(* IEC 61131-3 sources: daoli-st-library/DL_Base (part 12) *)

(* ---- FB_DL_EventCounter.st ---- *)
(*==============================================================================
 * 组件名称 (Component)  : FB_DL_EventCounter
 * 所属子库 (Sublibrary) : DL_Base
 * 当前版本 (Version)    : 1.0.1
 * 兼容性   (Platform)   : CODESYS 3.5 / TwinCAT 3 / 汇川 InoProShop / Machine Expert
 *                         仅依赖 Standard.library（R_TRIG），零厂商方言
 * 分类     (Category)   : 信号处理功能块（Function Block · 通用事件计数）
 * 功能简述 (Function)   : 双向事件计数器（DINT 域）。递增/递减脉冲沿独立
 *                         计数、预置装载、高/低阈值比较输出（每拍重算非锁
 *                         存）、回绕/饱和两种越界模式可选；双脉冲同拍抵消
 *                         置信息级、装载覆盖计数置信息级；参数非法故障锁存。
 *                         与 FC_DL_BitCount（位统计）、FB_DL_RuntimeMeter
 *                         （时间累计）职责分离，本块为通用事件计数。
 * 公约遵循 (Convention) : 0.1/R23 事件型，免首扫——计数由脉冲沿驱动，无
 *                         初始化/跟踪同步语义，不设 bInit。
 *                         0.2/R21 bFault 为显式排除信息级码的派生式；故障
 *                         码表逐条标注级别；信息级只进 uErrorId 不进报警链。
 *                         0.7/R15 故障级锁存仅解除路径（bReset 上升沿）清
 *                         码；信息级瞬时型每拍重算。
 *                         0.8 故障码段位 16#0001_xxxx（经 DL_Base VERSION.md
 *                         码表核对，0001_0101~0104 / 0001_0210 均未占用）：
 *                         【故障级】0001_0210 计数下限 ≥ 上限；
 *                         【信息级】0001_0101 双脉冲同拍抵消、0001_0102 装
 *                         载覆盖计数（bLoad 优先级最高，同拍覆盖计数脉冲）。
 * 红线自检 (Redline)    : R1 零全局变量表/外部变量引用 ✓｜R2 零物理 IO 地址 ✓
 *                         R3 纯 IEC 61131-3 ✓｜R4 越界钳位/回绕双模式 ✓
 *                         R5 全变量中英双语同行注释 ✓｜R7 三个边沿实例主体
 *                         最前部无条件刷新 ✓｜R8 越界常量化无魔法数 ✓
 * 设计要点 (Key notes)  : ① 双脉冲同拍到达：净变化 0，置信息级 0001_0101，
 *                           不计数（避免扫描时序歧义）；
 *                         ② 回绕语义：计数值越过 nMax → 回 nMin 继续（bWrap
 *                           =TRUE）；饱和语义：钳位在 nMax/nMin 并置溢出标志
 *                           一拍（bWrap=FALSE）；
 *                         ③ bLoad 上升沿优先级最高：同拍覆盖计数脉冲，置信
 *                           息级 0001_0102；
 *                         ④ bCompHigh = nCount >= nCompHigh、bCompLow =
 *                           nCount <= nCompLow，每拍重算非锁存（判据语义在
 *                           注释写死，防现场误解）；
 *                         ⑤ bOverflow/bUnderflow 为事件一拍脉冲，不锁存。
 * 开源溯源 (Origin)     : 来源标签 lgf-counter（RAW_NOTES_R7 S-1：LGF 库
 *                         CTU/CTUD 计数器族的功能语义域——双向计数、预置
 *                         装载、比较输出、回绕，公开文档，仅借鉴功能域语
 *                         义；实现、故障码与引脚契约 100% 本库独立设计，
 *                         clean-room 未复制源码）。
 * 验收向量 (Acceptance) :
 *   V1 增/减/抵消逐拍推演：单发 +1 → 1；再单发 -1 → 0；同拍双发 → 0 且
 *      信息级 0001_0101；
 *   V2 回绕跨上下限：nMin=0/nMax=9/bWrap=TRUE，nCount=9 时 +1 → 0 且
 *      bOverflow 一拍；nCount=0 时 -1 → 9 且 bUnderflow 一拍；
 *   V3 饱和钳位：bWrap=FALSE，nCount=9 时 +1 → 9（钳位）且 bOverflow 一拍；
 *   V4 预置装载：bLoad 沿 → nCount := nPreset=5；同拍 +1 脉冲被覆盖且信息
 *      级 0001_0102；
 *   V5 参数非法：nMin=10 > nMax=5 → 故障锁存 0001_0210，bFault=TRUE；
 *   V6 复位清零：bReset 沿 → 计数值=0、故障与信息码清零。
 * 修订历史 (Revision)   :
 *   2026-11-15  v1.0.0  首版入库（Round 07 · DL_Base LGF Counter 组开组）
 *   2026-11-15  v1.0.1  终审修复 2 处：① DINT 极值 +1/-1 回绕穿透饱和/回绕
 *                       判据（加算/减算改先判界后运算）；② 复位与计数脉冲
 *                       同拍时计数覆盖复位（复位拍最高优先，段 4 前置分支）
 *============================================================================*)
FUNCTION_BLOCK FB_DL_EventCounter
VAR_INPUT
    bCntUp     : BOOL;              // 递增计数脉冲（Count-up pulse），R_TRIG 上升沿 +1 / Count-up pulse, rising edge +1
    bCntDown   : BOOL;              // 递减计数脉冲（Count-down pulse），R_TRIG 上升沿 -1 / Count-down pulse, rising edge -1
    bLoad      : BOOL;              // 预置装载指令（Preset load），R_TRIG 上升沿把 nPreset 写入计数值 / Preset load edge writes nPreset into the count
    nPreset    : DINT;              // 预置值（Preset value）[-]，任意 DINT 域 / Preset value, any DINT value
    bWrap      : BOOL;              // 回绕模式使能（Wrap-around enable），TRUE=上溢回 nMin/nMax 循环；FALSE=饱和钳位 / TRUE = wrap to opposite limit, FALSE = saturate
    nMin       : DINT := -2147483648; // 计数下限（Count lower limit）[-]，默认 DINT 域下界（与 DL_CNT_DINT_MIN 一致）/ Lower limit, DINT minimum by default
    nMax       : DINT := 2147483647;  // 计数上限（Count upper limit）[-]，默认 DINT 域上界（与 DL_CNT_DINT_MAX 一致）/ Upper limit, DINT maximum by default
    nCompHigh  : DINT;              // 高阈值比较（High compare）[-]，bCompHigh 判据 nCount >= nCompHigh / High threshold for bCompHigh (greater-or-equal)
    nCompLow   : DINT;              // 低阈值比较（Low compare）[-]，bCompLow 判据 nCount <= nCompLow / Low threshold for bCompLow (less-or-equal)
    bReset     : BOOL;              // 上升沿复位故障与清零计数值（Reset edge clears fault and count）/ Rising edge resets fault and clears count
END_VAR
VAR_OUTPUT
    nCount      : DINT;             // 当前计数值（Current count）[-] / Current count value
    bCompHigh   : BOOL;             // 高阈值比较结果（High compare output），每拍重算 nCount >= nCompHigh 非锁存 / High compare, recomputed every scan, not latched
    bCompLow    : BOOL;             // 低阈值比较结果（Low compare output），每拍重算 nCount <= nCompLow 非锁存 / Low compare, recomputed every scan, not latched
    bOverflow   : BOOL;             // 上溢事件标志（Overflow event），本拍发生上溢置位一拍 / Overflow event, TRUE for one scan on overflow
    bUnderflow  : BOOL;             // 下溢事件标志（Underflow event），本拍发生下溢置位一拍 / Underflow event, TRUE for one scan on underflow
    bFault      : BOOL;             // 故障标志（Fault flag），显式排除信息级码（R21）/ Fault flag, info codes explicitly excluded
    uErrorId    : UDINT;            // 故障码（Error code），16#0001_xxxx 段，0=无故障 / Error code, family 16#0001_xxxx, 0 = none
END_VAR
VAR
    _fbTrigUp    : R_TRIG;          // 递增脉冲上升沿（Up pulse rising edge）/ Up pulse edge detector
    _fbTrigDown  : R_TRIG;          // 递减脉冲上升沿（Down pulse rising edge）/ Down pulse edge detector
    _fbTrigLoad  : R_TRIG;          // 装载指令上升沿（Load command rising edge）/ Load command edge detector
    _fbTrigReset : R_TRIG;          // 复位上升沿（Reset rising edge）/ Reset edge detector
    _bFaultLatch : BOOL;            // 故障锁存标志（Fault latch flag），仅 bReset 上升沿清除 / Fault latch, cleared only by reset edge
    _uErrorIdInt : UDINT;           // 内部故障级码寄存（Internal fault-level code register）/ Internal fault-level code register
    _uInfoCode   : UDINT;           // 本拍信息级码（Info code this cycle），瞬时型每拍重算 / Transient info code, recomputed each scan
    _bUpEdge     : BOOL;            // 本拍递增沿有效（Up edge active this scan）/ Up edge active this scan
    _bDownEdge   : BOOL;            // 本拍递减沿有效（Down edge active this scan）/ Down edge active this scan
    _bLoadEdge   : BOOL;            // 本拍装载沿有效（Load edge active this scan）/ Load edge active this scan
    _nWork       : DINT;            // 计数运算工作副本（Working copy of count）[-] / Working copy for arithmetic
END_VAR
VAR CONSTANT
    DL_CNT_DINT_MIN : DINT := -2147483648; // DINT 域下界（DINT lower bound）/ DINT lower bound
    DL_CNT_DINT_MAX : DINT := 2147483647;  // DINT 域上界（DINT upper bound）/ DINT upper bound
END_VAR

// ============================================================================
// 段 1｜边沿实例无条件周期刷新（R7/0.5：严禁置于 IF/CASE 分支内）
//      Unconditional per-cycle refresh of all edge instances (R7/0.5)
// ============================================================================
_fbTrigUp(CLK    := bCntUp);
_fbTrigDown(CLK  := bCntDown);
_fbTrigLoad(CLK  := bLoad);
_fbTrigReset(CLK := bReset);
_bUpEdge   := _fbTrigUp.Q;        // 本拍递增沿（Up edge this scan）
_bDownEdge := _fbTrigDown.Q;      // 本拍递减沿（Down edge this scan）
_bLoadEdge := _fbTrigLoad.Q;      // 本拍装载沿（Load edge this scan）

// ============================================================================
// 段 2｜信息级码预清零 + 复位路径（R15：锁存型故障只在解除路径清码）
//      Info code preset zero + reset path (R15: latched fault cleared in release path only)
// ============================================================================
_uInfoCode := 0;                  // 信息级瞬时型每拍重算（Transient info recomputed each scan）
bOverflow  := FALSE;              // 事件标志每拍预清零，由段 4 事件置位一拍（Event flags preset FALSE, set one scan by stage 4）
bUnderflow := FALSE;              // 事件标志每拍预清零（Event flag preset FALSE）

IF _fbTrigReset.Q THEN
    _nWork      := 0;             // 计数值清零（Count cleared）
    _bFaultLatch := FALSE;        // 故障锁存解除（Fault latch released）
    _uErrorIdInt := 16#0000_0000; // 故障码清零（Fault code cleared）
END_IF

// ============================================================================
// 段 3｜参数防御：nMin >= nMax → 故障锁存（故障级，锁存期间计数值冻结）
//      Parameter guard: nMin >= nMax latches a fault-level error, count frozen
// ============================================================================
IF nMin >= nMax THEN
    _bFaultLatch := TRUE;                 // 参数非法故障锁存（Invalid limit latch）
    _uErrorIdInt := 16#0001_0210;         // 0001_0210 计数下限 ≥ 上限【故障级】/ Lower limit >= upper limit, fault level
ELSE

    // ========================================================================
    // 段 4｜计数主逻辑：装载优先 → 双脉冲抵消 → 单向计数与越界处理
    //      Counting main logic: load first, dual-pulse cancellation, then counting
    // ========================================================================
    IF _fbTrigReset.Q THEN
        _nWork := 0;                    // 复位拍最高优先：同拍计数/装载脉冲被复位覆盖（复位-计数同拍冲突修复）/ Reset scan top priority, pulses overridden
    ELSIF _bLoadEdge THEN
        _nWork := nPreset;                // 装载优先级最高：预置值直接写入（Load has top priority）
        IF _bUpEdge OR _bDownEdge THEN
            _uInfoCode := 16#0001_0102;   // 0001_0102 装载覆盖计数【信息级】/ Load overrides counting pulses, info level
        END_IF
    ELSIF _bUpEdge AND _bDownEdge THEN
        _uInfoCode := 16#0001_0101;     // 0001_0101 双脉冲同拍抵消【信息级】，净变化 0 / Dual pulses cancel, net zero, info level
    ELSIF _bUpEdge THEN
        // 先判界再加算：nCount 已达 nMax 直接走越界语义，杜绝 DINT 极值 +1
        // 回绕穿透（nCount=DINT_MAX 时 +1 回绕为负、>nMax 判据失效）
        // Boundary pre-check before increment: DINT-max +1 wrap cannot bypass the verdict
        IF nCount >= nMax THEN
            IF bWrap THEN
                _nWork := nMin;         // 回绕语义：越过上限回下限（Wrap: above max falls back to min）
            ELSE
                _nWork := nMax;         // 饱和语义：钳位在上限（Saturate at max）
            END_IF
            bOverflow := TRUE;          // 上溢事件一拍脉冲（Overflow event, one scan）
        ELSE
            _nWork := nCount + 1;       // 递增一步（Increment one step, pre-guarded no-overflow）
        END_IF
    ELSIF _bDownEdge THEN
        // 先判界再减算：对称防御 DINT 极值 −1 回绕穿透（Mirror of the increment guard）
        IF nCount <= nMin THEN
            IF bWrap THEN
                _nWork := nMax;         // 回绕语义：越过下限回上限（Wrap: below min jumps to max）
            ELSE
                _nWork := nMin;         // 饱和语义：钳位在下限（Saturate at min）
            END_IF
            bUnderflow := TRUE;         // 下溢事件一拍脉冲（Underflow event, one scan）
        ELSE
            _nWork := nCount - 1;       // 递减一步（Decrement one step, pre-guarded no-overflow）
        END_IF
    ELSE
        _nWork := nCount;               // 无事件保持计数值（No event, hold count）
    END_IF
    nCount := _nWork;                   // 计数值单点出口（Single outlet for the count）
END_IF

// ============================================================================
// 段 5｜输出推导：比较输出每拍重算、溢出标志由段 4 置位本拍后自然回落
//      Output derivation: compare outputs recomputed each scan, event flags one-shot
// ============================================================================
bCompHigh := (nCount >= nCompHigh);   // 高阈值判据（High compare: greater-or-equal）
bCompLow  := (nCount <= nCompLow);    // 低阈值判据（Low compare: less-or-equal）

IF _fbTrigReset.Q THEN
    bOverflow  := FALSE;              // 复位拍清事件标志（Event flags cleared on reset scan）
    bUnderflow := FALSE;
END_IF

IF _bFaultLatch THEN
    nCount := 0;                      // 故障期计数值输出安全零（Safe zero while latched）
END_IF

// ============================================================================
// 段 6｜bFault/uErrorId 出口（R21：bFault 显式排除信息级；无故障级锁存时
//       uErrorId 透出本拍信息级码）
//      Outlets: bFault excludes info codes (R21); uErrorId shows info code when no fault
// ============================================================================
bFault := _bFaultLatch;               // 故障级派生式（Fault-level derived form）
IF _bFaultLatch THEN
    uErrorId := _uErrorIdInt;         // 故障级码优先透出（Fault-level code has priority）
ELSE
    uErrorId := _uInfoCode;           // 无故障时透出本拍信息级码（Transient info code when no fault）
END_IF
END_FUNCTION_BLOCK

(* ---- FB_DL_ExtendedTimer.st ---- *)
(*==============================================================================
 * 组件名称 (Component)  : FB_DL_ExtendedTimer
 * 所属子库 (Sublibrary) : DL_Base
 * 当前版本 (Version)    : 1.0.0
 * 兼容性   (Platform)   : CODESYS 3.5 / TwinCAT 3 / 汇川 InoProShop / Machine Expert
 *                         仅依赖 Standard.library（TON / R_TRIG / F_TRIG），零厂商方言
 * 功能描述 (Function)   : 四模式工业定时器，一个实例覆盖通电延时 / 断电延时 / 单脉冲 /
 *                         保持型累加四种现场时序需求，消除"同一延时逻辑在项目里
 *                         散落四种实现、改造时漏改某处"的维护风险。
 *                         保持型累加模式补足标准库空白：输入断开时进度保留，
 *                         只有显式复位才清零，累加采用相位定时器差值累加而非直读已计时值。
 *                         运行中切换模式立即作废当前计时（操作语义，不产生故障码）。
 * 开源溯源 (Origin)     : 原创实现。四模式语义依据 IEC 61131-3 标准 TON/TOF/TP 定义，
 *                         保持型累加模式参照 AB / Omron 生态的 RTO 行为定义；
 *                         全部代码为本库独立重构，未复制任何厂商或开源库源码。
 * 本文件内含       : TYPE  E_DL_TimerMode（配套枚举，归属 DL_Base）
 *                    TYPE  E_DL_ExtTimerState（配套枚举，归属 DL_Base）
 *                    FB    FB_DL_ExtendedTimer
 * 依赖     (Depends)    : 无 DL_ 内部依赖；Standard.library: TON / R_TRIG / F_TRIG
 * 红线自检 (Redline)    : R1 ✓ 禁用全局存储与物理寻址 ｜ R2 ✓ 无地址直写
 *                         R3 ✓ 纯 IEC 61131-3 ｜ R4 ✓ 预设钳位 + 剩余时间负值钳位 + 差分累加防倒退
 *                         R5 ✓ 全变量中英双语同行注释 ｜ R6 ✓ 四态 ENUM + CASE + ELSE 兜底
 *                         R7 ✓ 三实例主体最前部无条件刷新（本组件核心考点）
 *                         R8 ✓ 预设上限、零值判据全常量化
 *
 * 【四模式输出语义表 / Four-mode output semantics（边界 B2，手册原样收录）】
 *   通电延时：输入 TRUE 满 PT 后输出 TRUE；输入 FALSE 立即输出 FALSE 且已计时清零。
 *   断电延时：输入 TRUE 期间输出 TRUE；输入变 FALSE 后输出保持 TRUE 并计时，
 *             满 PT 才复位为 FALSE；输入提前恢复 TRUE 则计时作废。
 *   单脉冲  ：输入上升沿触发，输出 TRUE 持续 PT 时长；期间输入变 FALSE 不中断；
 *             新上升沿重触发并从零重新计时。
 *   保持型  ：输入 TRUE 时累加计时，输入 FALSE 时进度保留不清零；
 *             累计达 PT 后输出 TRUE 且不再受输入影响，仅复位可清零。
 *
 * 【模式切换即计时作废 / Mode switch voids the timing（边界 B4）】
 *   运行中改写模式会立即中止当前计时、清零累加并回到待机态，
 *   这是操作语义而不是故障，因此不产生任何故障码（手册须写明）。
 *
 * 修订历史 (Revision)   :
 *   2026-11-14  v1.0.0  首版入库（Phase 1 第二轮 · Level 0 批次 B）
 *============================================================================*)

(*-----------------------------------------------------------------------------
 * 枚举: E_DL_TimerMode（归属 DL_Base，与 FB_DL_ExtendedTimer 同文件）
 * 含义: 定时器工作模式。数值与现场惯用编号一致，便于 HMI 配方直接映射。
 *----------------------------------------------------------------------------*)
TYPE E_DL_TimerMode :
(
    eTon := 0,    // 通电延时：输入保持 TRUE 满 PT 后输出 TRUE / On-delay, output TRUE after PT of TRUE input
    eTof := 1,    // 断电延时：输入变 FALSE 后延时 PT 再复位输出 / Off-delay, output drops PT after the input falls
    eTp  := 2,    // 单脉冲：上升沿触发 PT 时长脉冲，可重触发 / Pulse, retriggerable on each rising edge
    eRto := 3     // 保持型累加：输入 TRUE 累加，断开保持进度，仅复位清零 / Retentive on-delay, reset only
);
END_TYPE

(*-----------------------------------------------------------------------------
 * 枚举: E_DL_ExtTimerState（归属 DL_Base，与 FB_DL_ExtendedTimer 同文件）
 * 含义: 定时器主状态。数值步长留空位便于后续插态而不破坏已有工程。
 *----------------------------------------------------------------------------*)
TYPE E_DL_ExtTimerState :
(
    eIdle   := 0,     // 待机：输出为当前模式的待机值 / Idle, output at the mode rest value
    eTiming := 10,    // 计时进行中 / Timing in progress
    eDone   := 20,    // 完成：输出保持 / Done, output held
    eFault  := 99     // 故障锁定：需复位清除 / Fault latched, cleared by reset
);
END_TYPE

FUNCTION_BLOCK FB_DL_ExtendedTimer
VAR_INPUT
    bIn      : BOOL;                        // 输入信号（电平语义）/ Input signal, level semantics
    eMode    : E_DL_TimerMode := eTon;      // 工作模式 / Operating mode
    tPreset  : TIME := T#10S;               // 预设时间 [ms]，合法域 0 至上限 / Preset time [ms], valid range up to the clamp
    bReset   : BOOL;                        // 上升沿：清零累加与故障 / Rising edge: clear the accumulation and the fault
END_VAR
VAR_OUTPUT
    bQ         : BOOL;    // 输出，语义随模式（见头注释语义表）/ Output, semantics per mode, see the header table
    bTiming    : BOOL;    // 计时进行中标志 / Timing in progress flag
    tElapsed   : TIME;    // 当前模式已计时 [ms]，保持型为累计值 / Elapsed time [ms], accumulated in retentive mode
    tRemaining : TIME;    // 距完成剩余 [ms]，完成或待机为 0 / Remaining time [ms], zero when done or idle
    uErrorId   : UDINT;   // 故障码，0 = 无故障 / Error code, 0 = no error
END_VAR
VAR
    fbTrigRise  : R_TRIG;                 // 输入上升沿检测实例 / Input rising edge detector instance
    fbTrigFall  : F_TRIG;                 // 输入下降沿检测实例 / Input falling edge detector instance
    fbTrigReset : R_TRIG;                 // 复位上升沿检测实例 / Reset rising edge detector instance
    fbTonPhase  : TON;                    // 相位计时器，四模式共用 / Phase timer shared by all four modes
    eState      : E_DL_ExtTimerState;     // 主状态机 / Main state machine
    tAccum      : TIME;                   // 保持型累计时间 [ms] / Retentive accumulated time [ms]
    eLastMode   : E_DL_TimerMode;         // 上周期模式，用于变更检测 / Previous mode for change detection
    tPresetEff  : TIME;                   // 钳位后的预设时间 [ms] / Clamped preset time [ms]
    tTonPt      : TIME;                   // 相位定时器当前预设 [ms] / Current preset of the phase timer [ms]
    tEtPrev     : TIME;                   // 上周期相位定时器已计时 [ms]，差分累加用 / Previous ET for delta accumulation [ms]
    tDelta      : TIME;                   // 本周期已计时增量 [ms] / ET increment of this scan [ms]
    bTonIn      : BOOL;                   // 相位定时器输入（先推导后喂入）/ Phase timer input, derived first then fed
    bModeBad    : BOOL;                   // 模式枚举越界标志 / Mode enum out-of-domain flag
    bPresetBad  : BOOL;                   // 预设时间越界标志 / Preset out-of-range flag
    bPresetZero : BOOL;                   // 预设为零标志（立即完成）/ Zero preset flag, complete immediately
    bRtoDone    : BOOL;                   // 保持型累加已达标（锁存）/ Retentive accumulation reached the preset, latched
    bTofArmed   : BOOL;                   // 断电延时的延时阶段已建立 / Off-delay hold phase armed
    bTpRun      : BOOL;                   // 单脉冲进行中 / Single pulse running
    bHoldOn     : BOOL;                   // 本周期强制定时器停计（复位/换模式/故障）/ Force the timer off this scan
END_VAR
VAR CONSTANT
    DL_TIMER_PRESET_MAX : TIME := T#12H;  // 预设时间上限钳位 [h] / Preset clamp [h]
END_VAR

(*------------------------------------------------------------------------------
 * 段 1｜无条件刷新区（红线 R7 / 边界 B1）：三个实例严禁进入任何 IF / CASE 分支
 *      Unconditional refresh zone: no instance call inside IF / CASE
 *      IN 与 PT 均由"状态 + 输入"先行推导成普通量，实例调用本身保持无条件
 *      IN and PT are derived into plain values first, the calls stay unconditional
 *-----------------------------------------------------------------------------*)
fbTrigRise(CLK  := bIn);
fbTrigFall(CLK  := bIn);
fbTrigReset(CLK := bReset);

(*------------------------------------------------------------------------------
 * 段 2｜预设钳位（边界 B3）：超上限钳到上限并告警，但计时继续不中断
 *      Preset clamping: clamp and warn, but keep timing without interruption
 *-----------------------------------------------------------------------------*)
bPresetBad := FALSE;

IF tPreset > DL_TIMER_PRESET_MAX THEN
    tPresetEff := DL_TIMER_PRESET_MAX;
    bPresetBad := TRUE;
ELSIF tPreset < T#0S THEN
    tPresetEff := T#0S;
    bPresetBad := TRUE;
ELSE
    tPresetEff := tPreset;
END_IF

bPresetZero := (tPresetEff <= T#0S);

(*------------------------------------------------------------------------------
 * 段 3｜模式合法性（边界 B7）：枚举被强制写入域外值时直接进故障态
 *      Mode validity: an out-of-domain enum drives the state machine to fault
 *-----------------------------------------------------------------------------*)
bModeBad := NOT ((eMode = eTon) OR (eMode = eTof) OR (eMode = eTp) OR (eMode = eRto));

(*------------------------------------------------------------------------------
 * 段 4｜运行中模式切换（边界 B4）：立即中止计时、清零累加，不产生故障码
 *      Mode switch while running: abort the timing and clear the accumulation, no error
 *      本周期强制定时器停计，让相位定时器在下一周期从零重新起算
 *      The timer is forced off this scan so it restarts from zero next scan
 *-----------------------------------------------------------------------------*)
bHoldOn := FALSE;

IF eMode <> eLastMode THEN
    eLastMode := eMode;
    eState    := eIdle;
    tAccum    := T#0S;
    tEtPrev   := T#0S;
    bRtoDone  := FALSE;
    bTofArmed := FALSE;
    bTpRun    := FALSE;
    bHoldOn   := TRUE;
END_IF

(*------------------------------------------------------------------------------
 * 段 5｜相位定时器输入推导（边界 B2）：先算成 BOOL，再喂给实例
 *      Phase timer input derivation: compute the BOOL first, then feed the instance
 *      四种模式对"何时计时"的要求完全不同，统一收敛到一个推导段便于审阅
 *      All four modes converge here so the timing condition is reviewed in one place
 *-----------------------------------------------------------------------------*)
bTonIn := FALSE;
tTonPt := tPresetEff;

IF bModeBad THEN
    bTonIn := FALSE;
ELSIF eMode = eTon THEN
    (* 通电延时：输入为 TRUE 即计时 *)
    (* On-delay: time while the input is TRUE *)
    bTonIn := bIn;
ELSIF eMode = eTof THEN
    (* 断电延时：输入为 FALSE 即计时（输入 TRUE 时 ET 被清零） *)
    (* Off-delay: time while the input is FALSE, a TRUE input clears ET *)
    bTonIn := NOT bIn;
ELSIF eMode = eTp THEN
    (* 单脉冲：上升沿当周期强制停计一拍，使 ET 清零后重新计时（可重触发） *)
    (* Pulse: the rising scan forces one off-scan so ET restarts from zero *)
    bTonIn := bTpRun AND (NOT fbTrigRise.Q);
ELSE
    (* 保持型：输入 TRUE 且未达标时计时 *)
    (* Retentive: time while the input is TRUE and the preset is not yet reached *)
    bTonIn := bIn AND (NOT bRtoDone);
END_IF

(*------------------------------------------------------------------------------
 * 段 6｜相位定时器无条件刷新（红线 R7）：全组件唯一一次调用
 *      Single unconditional call of the phase timer
 *      复位 / 换模式 / 故障 / 禁用当周期统一断开 IN，ET 由标准语义自动清零
 *      Reset, mode switch and fault all drop IN so the standard semantics clear ET
 *-----------------------------------------------------------------------------*)
fbTonPhase(IN := bTonIn AND (NOT bHoldOn) AND (NOT fbTrigReset.Q) AND (NOT bModeBad) AND (eState <> eFault),
           PT := tTonPt);

(*------------------------------------------------------------------------------
 * 段 7｜保持型差分累加（边界 B5）：把 ET 的增量并入累计，禁止直读 ET 当累计值
 *      Retentive delta accumulation: fold the ET increment into the accumulator
 *      ET 在输入断开时会被标准定时器清零，若直读 ET 当累计值，进度当场丢失
 *      ET is cleared when the input drops, reading it directly would lose the progress
 *      增量为负说明定时器刚被清零，忽略即可，累计值因此只增不减
 *      A negative delta means the timer just reset, ignoring it keeps the total monotonic
 *-----------------------------------------------------------------------------*)
IF (eMode = eRto) AND (NOT bModeBad) AND (NOT bRtoDone) THEN
    tDelta := fbTonPhase.ET - tEtPrev;
    IF tDelta > T#0S THEN
        tAccum := tAccum + tDelta;
        IF tAccum >= tPresetEff THEN
            tAccum   := tPresetEff;
            bRtoDone := TRUE;
        END_IF
    END_IF
END_IF

tEtPrev := fbTonPhase.ET;

(*------------------------------------------------------------------------------
 * 段 8｜复位语义（边界 B6）：保持型唯一清零路径，同时清故障与全部模式标志
 *      Reset: the only clearing path of the retentive accumulator
 *-----------------------------------------------------------------------------*)
IF fbTrigReset.Q THEN
    eState    := eIdle;
    tAccum    := T#0S;
    tEtPrev   := T#0S;
    bRtoDone  := FALSE;
    bTofArmed := FALSE;
    bTpRun    := FALSE;
    bPresetBad := FALSE;
    uErrorId  := 16#0000_0000;
ELSE

    (*--------------------------------------------------------------------------
     * 段 9｜主状态机（红线 R6）：ENUM + CASE + ELSE 兜底
     *      Main state machine with the mandatory ELSE fallback
     *-------------------------------------------------------------------------*)
    IF bModeBad THEN
        eState := eFault;
    ELSE
        CASE eState OF

            eIdle:
                (* 待机态：按模式等待各自的启动事件 *)
                (* Idle: wait for the mode-specific start event *)
                IF eMode = eTon THEN
                    (* 预设为零时立即完成，不占一个扫描周期的启动延迟 *)
                    (* A zero preset completes immediately, no start-up scan delay *)
                    IF bIn AND bPresetZero THEN
                        eState := eDone;
                    ELSIF bIn THEN
                        eState := eTiming;
                    END_IF
                ELSIF eMode = eTof THEN
                    IF bIn THEN
                        bTofArmed := TRUE;
                        eState    := eDone;
                    END_IF
                ELSIF eMode = eTp THEN
                    IF fbTrigRise.Q THEN
                        bTpRun := TRUE;
                        eState := eTiming;
                    END_IF
                ELSE
                    (* 保持型：已达标或输入到来均可启动；进度保留在 tAccum *)
                    (* Retentive: resume from the retained accumulation *)
                    IF bRtoDone THEN
                        eState := eDone;
                    ELSIF bIn AND bPresetZero THEN
                        bRtoDone := TRUE;
                        eState   := eDone;
                    ELSIF bIn THEN
                        eState := eTiming;
                    END_IF
                END_IF

            eTiming:
                IF eMode = eTon THEN
                    (* 输入掉电立即回待机，输出与已计时一并清零（语义表第一行） *)
                    (* Input falling returns to idle and clears the elapsed time *)
                    IF NOT bIn THEN
                        eState := eIdle;
                    ELSIF fbTonPhase.Q THEN
                        eState := eDone;
                    END_IF
                ELSIF eMode = eTof THEN
                    (* 输入恢复：延时作废回完成态；延时到期：回待机 *)
                    (* Input recovered voids the delay, expiry returns to idle *)
                    IF bIn THEN
                        eState := eDone;
                    ELSIF fbTonPhase.Q THEN
                        bTofArmed := FALSE;
                        eState    := eIdle;
                    END_IF
                ELSIF eMode = eTp THEN
                    (* 脉冲期满：结束脉冲；期间输入变化不打断，新上升沿由段 5 重触发 *)
                    (* Pulse expiry ends the pulse, a new rising edge retriggers via stage 5 *)
                    IF fbTonPhase.Q THEN
                        bTpRun := FALSE;
                        eState := eDone;
                    END_IF
                ELSE
                    (* 保持型：达标锁存；输入断开回待机但累计值保留 *)
                    (* Retentive: latch on done, an input drop keeps the accumulation *)
                    IF bRtoDone THEN
                        eState := eDone;
                    ELSIF NOT bIn THEN
                        eState := eIdle;
                    END_IF
                END_IF

            eDone:
                IF eMode = eTon THEN
                    IF NOT bIn THEN
                        eState := eIdle;
                    END_IF
                ELSIF eMode = eTof THEN
                    (* 输入断开即进入延时阶段 *)
                    (* An input drop starts the off-delay phase *)
                    IF NOT bIn THEN
                        eState := eTiming;
                    END_IF
                ELSIF eMode = eTp THEN
                    (* 脉冲结束后等待下一次上升沿 *)
                    (* Wait for the next rising edge after the pulse finished *)
                    IF fbTrigRise.Q THEN
                        bTpRun := TRUE;
                        eState := eTiming;
                    END_IF
                ELSE
                    (* 保持型：达标后锁存，仅段 8 的复位可解除 *)
                    (* Retentive: latched after done, only the reset in stage 8 clears it *)
                    eState := eDone;
                END_IF

            eFault:
                (* 故障锁存：输出由段 10 强制 FALSE，等待复位 *)
                (* Fault latched: stage 10 forces the output FALSE until reset *)
                eState := eFault;

            ELSE
                (* 非法状态拦截：转故障并上报，不做隐式恢复 *)
                (* Illegal state interception: go to fault and report, no implicit recovery *)
                eState := eFault;

        END_CASE;
    END_IF
END_IF

(*------------------------------------------------------------------------------
 * 段 10｜输出单一出口（边界 B8 / P-05）：三个输出只在此处统一赋值一次
 *      Single output outlet: the three outputs are written exactly once here
 *      分支内部只改状态与标志，不直接写输出，避免同一输出在多处赋值产生竞态
 *      Branches only change state and flags, never the outputs, to avoid races
 *-----------------------------------------------------------------------------*)
CASE eMode OF
    eTon:
        bQ := (eState = eDone);
    eTof:
        (* 输入 TRUE 期间与延时保持期间均输出 TRUE *)
        (* TRUE while the input is TRUE and during the off-delay hold *)
        bQ := (eState = eTiming) OR (eState = eDone);
    eTp:
        bQ := (eState = eTiming);
    eRto:
        bQ := (eState = eDone);
    ELSE
        bQ := FALSE;
END_CASE;

IF eState = eFault THEN
    bQ := FALSE;
END_IF

IF eMode = eRto THEN
    (* 保持型输出累计值：输入断开后进度仍可见，这是该模式的存在意义 *)
    (* The retentive mode reports the accumulation so the progress stays visible *)
    tElapsed := tAccum;
ELSE
    IF (eState = eIdle) OR (eState = eFault) THEN
        tElapsed := T#0S;
    ELSE
        tElapsed := fbTonPhase.ET;
    END_IF
END_IF

(* 剩余时间负值钳位（边界 B9）：换算与时序竞态都可能产生负差，一律钳到零 *)
(* Remaining time clamp: rounding and timing races can go negative, clamp to zero *)
IF tElapsed >= tPresetEff THEN
    tRemaining := T#0S;
ELSE
    tRemaining := tPresetEff - tElapsed;
END_IF

bTiming := (eState = eTiming);

(*------------------------------------------------------------------------------
 * 段 11｜故障码汇总：模式越界 > 非法状态 > 预设钳位
 *      Error aggregation: mode out-of-domain, illegal state, then preset clamp
 *-----------------------------------------------------------------------------*)
IF bModeBad THEN
    uErrorId := 16#0001_000E;
ELSIF eState = eFault THEN
    uErrorId := 16#0001_0005;
ELSIF bPresetBad THEN
    uErrorId := 16#0001_0001;
ELSE
    uErrorId := 16#0000_0000;
END_IF
END_FUNCTION_BLOCK

(* ---- FB_DL_FirstOutLatch.st ---- *)
(*
    FB_DL_FirstOutLatch —— 多源故障首出锁存
    ------------------------------------------------------------------
    分类      : DL_Base / Signal
    前缀      : FB_DL_
    版本      : 1.0.0
    溯源      : T2-8 ISA-18.2 公开的「首出 / 确认 / 锁存」生命周期语义；
                本库 FB_DL_PortDiagAggregator 首出三律（最小序号仲裁）同口径复用。
                只借公开首出语义与仲裁次序，不借任何实现代码行；clean-room 重写，
                未复制任何闭源厂商源码，参考实现仅限 MIT/Apache 许可
    平台      : 纯 IEC 61131-3，CODESYS V3.5+ / TwinCAT 3 / InoProShop 通用
    作者      : 道莅代码库 · PLC编程专家（R18）
    ------------------------------------------------------------------
    功能说明  : 16 路故障源并行输入，首个到来的源被锁存为唯一「首出原因」，后续源
                不得覆盖；bReset 上升沿清锁存且当拍不重新锁存（防复位自杀）；
                同拍多源按源序号最小仲裁，与库内首出三律同一口径，避免两套规则；
                uSrcCount 越界时不索引数组、全输出回安全值；
                bAnyFault / uFaultWord 为组合量（每拍重算不锁存），
                bLatched / uFirstIdx 为锁存量（仅复位或失能清除）。
    错误码    : 16#0001_0235 同拍多源故障，已按源序号最小仲裁为唯一首出——信息级，正常防御
                16#0001_0236 预留禁用（信息级，不得挪用）
                16#0001_0306 源数量参数越界（uSrcCount 不在 1~16）——故障级，本拍不锁存
                16#0001_0307 预留禁用（故障级，不得挪用）
                16#0001_0308 预留禁用（故障级，不得挪用）
    码位总账  : 16#0001_0235 用 / 16#0001_0236 预留 ｜ 16#0001_0306 用 / 16#0001_0307 预留 / 16#0001_0308 预留
    状态机    : 无 CASE，锁存由单比特保持（bLatchedInt），非法状态不可能出现，故以本节说明替代 ELSE 兜底
    采样约定  : bReset 的上升沿由 R_TRIG 在本体首部无条件刷新，绝不放入条件分支；
                本件无时间量参与，仲裁结果与任务周期无关，一个任务周期即完成一次仲裁。
    修订记录  : 2026-11-16 v1.0.0 首次入库（R18）
*)
FUNCTION_BLOCK FB_DL_FirstOutLatch
VAR_INPUT
    bEnable   : BOOL;                          // 使能，FALSE 清锁存并冻结仲裁 / enable, FALSE clears the latch and freezes arbitration
    bReset    : BOOL;                          // 复位，上升沿清首出锁存且当拍不重新锁存 / reset, rising edge clears the first-out latch and does not re-latch this cycle
    aSrcFault : ARRAY[0..15] OF BOOL;          // 16 路故障源，索引即优先级 0 最高 [路] / 16 fault sources, index is priority, 0 highest [ch]
    uSrcCount : UINT := 16;                    // 有效源数 [路]，范围 1~16 / valid source count [ch], range 1~16
END_VAR
VAR_OUTPUT
    bAnyFault : BOOL;                          // 任一源故障，组合值不锁存 / any source fault, combination value not latched
    bLatched  : BOOL;                          // 首出已被锁存 / first-out latched
    uFirstIdx : UINT;                          // 首出源序号 0~15，未锁存时为哨兵 16#FFFF / first-out index 0~15, sentinel 16#FFFF when not latched
    uFaultWord: WORD;                          // 当拍故障位图，bit0 = 源 0 [位图] / current fault bitmap, bit0 = source 0 [bitmap]
    eErr      : UDINT;                         // 错误码，0=正常 / error id, 0=ok
    bError    : BOOL;                          // 故障标志，eErr 为故障级时 TRUE / error flag, TRUE on fault-level eErr
END_VAR
VAR
    fbTrigReset : R_TRIG;                      // 复位上升沿检测实例，本体首部无条件刷新 / reset rising edge instance, refreshed unconditionally at body top
    uIdx        : UINT;                        // 源扫描游标 [路] / source scan cursor [ch]
    bAny        : BOOL;                        // 本拍存在故障源的中间标志 / intermediate flag, any source active this cycle
    bInit       : BOOL := FALSE;               // 首扫标志，初值 FALSE，判据 NOT bInit / first-scan flag, initial FALSE, tested with NOT
    bLatchedInt : BOOL;                        // 内部首出锁存位 / internal first-out latch bit
    uFirstInt   : UINT := 16#FFFF;             // 内部首出序号寄存，初值为哨兵 / internal first-out index register, initialised to the sentinel
    uActCnt     : UINT;                        // 本拍有效故障源计数，用于多源仲裁提示 [路] / active source count this cycle, used for the arbitration hint [ch]
END_VAR
VAR CONSTANT
    DL_FIRSTOUT_SRC_MAX : UINT := 16;          // 源上限 [路] / source upper bound [ch]
    DL_FIRSTOUT_NONE    : UINT := 16#FFFF;     // 无首出哨兵 [无量纲] / no-first-out sentinel [dimensionless]
    DL_FIRSTOUT_BIT_MAX : UINT := 15;          // 位图最高位号 [位] / highest bitmap index [bit]
    DL_FIRSTOUT_BIT0    : WORD := 16#0001;     // 位图最低位掩码 [位图] / least significant bitmap mask [bitmap]
END_VAR

// 段 1｜边沿实例无条件周期刷新（红线：严禁放入条件分支）/ segment 1, unconditional edge refresh
fbTrigReset(CLK := bReset);

// 段 2｜输出与中间量预置：组合量每拍重算，锁存量由内部位承载 / segment 2, preset outputs and temporaries
bAnyFault := FALSE;                            // 组合量先按无故障预置 / preset no fault on the combination output
uFaultWord := 0;                               // 位图先清零 / clear the bitmap
eErr := 0;                                     // 预置无错误 / preset no error
bError := FALSE;                               // 预置无故障标志 / preset no fault flag
bAny := FALSE;                                 // 中间标志清零 / clear the intermediate flag
uActCnt := 0;                                  // 有效源计数清零 / clear the active source count

// 段 3｜首扫初始化（唯一合法范式：初值 FALSE，判据 NOT bInit）/ segment 3, first-scan initialisation
IF NOT bInit THEN
    bLatchedInt := FALSE;                      // 首扫不留锁存 / no latch survives the first scan
    uFirstInt := DL_FIRSTOUT_NONE;             // 首出序号回哨兵 / first-out index back to the sentinel
    bInit := TRUE;                             // 首扫只做一次 / first scan runs once only
END_IF

// 段 4｜使能闸：失能清锁存并冻结，不索引数组 / segment 4, enable gate clears the latch and freezes
IF NOT bEnable THEN
    bLatchedInt := FALSE;                      // 清锁存位 / clear the latch bit
    uFirstInt := DL_FIRSTOUT_NONE;             // 清首出序号 / clear the first-out index
    bLatched := FALSE;                         // 对外锁存输出复位 / reset the latched output
    uFirstIdx := DL_FIRSTOUT_NONE;             // 对外序号回哨兵 / reset the index output to the sentinel
    RETURN;                                    // 失能即出口，本拍不仲裁 / disabled is the exit, no arbitration this cycle
END_IF

// 段 5｜源数量参数闸：越界即故障级，全输出回安全值且绝不索引数组 / segment 5, source count gate
IF (uSrcCount < 1) OR (uSrcCount > DL_FIRSTOUT_SRC_MAX) THEN
    eErr := 16#0001_0306;                      // 源数量越界故障码 / source count out of range fault id
    bError := TRUE;                            // 置故障标志 / raise the error flag
    bLatched := FALSE;                         // 锁存输出回安全值 / latched output to the safe value
    uFirstIdx := DL_FIRSTOUT_NONE;             // 序号输出回哨兵 / index output to the sentinel
    bLatchedInt := FALSE;                      // 内部锁存位清除 / clear the internal latch bit
    uFirstInt := DL_FIRSTOUT_NONE;             // 内部序号清除 / clear the internal index
    RETURN;                                    // 故障级提前返回 / early return on fault
END_IF

// 段 6｜组合扫描：位图与有效源计数（索引上界已由段 5 保证，位号不超过 15）/ segment 6, combination scan
FOR uIdx := 0 TO uSrcCount - 1 DO
    IF aSrcFault[uIdx] THEN
        bAny := TRUE;                          // 至少一源动作 / at least one source is active
        uActCnt := uActCnt + 1;                // 累加有效源数 / accumulate the active source count
        uFaultWord := uFaultWord OR SHL(DL_FIRSTOUT_BIT0, uIdx); // 置对应位，uIdx 不超过 15 故移位安全 / set the bit, uIdx never exceeds 15 so the shift is safe
    END_IF
END_FOR
bAnyFault := bAny;                             // 组合量对外输出 / publish the combination value

// 段 7｜复位沿优先于锁存（防自杀）：复位拍只清不锁 / segment 7, reset edge has priority over latching
IF fbTrigReset.Q THEN
    bLatchedInt := FALSE;                      // 复位清锁存 / reset clears the latch
    uFirstInt := DL_FIRSTOUT_NONE;             // 复位清序号 / reset clears the index
ELSIF (NOT bLatchedInt) AND bAny THEN
    FOR uIdx := 0 TO uSrcCount - 1 DO
        IF (uFirstInt = DL_FIRSTOUT_NONE) AND aSrcFault[uIdx] THEN
            uFirstInt := uIdx;                 // 只记第一个为真的源，索引最小即优先级最高 / record only the first active source, lowest index wins
        END_IF
    END_FOR
    bLatchedInt := TRUE;                       // 锁定首出 / latch the first-out source
    IF uActCnt > 1 THEN
        eErr := 16#0001_0235;                  // 同拍多源，已按最小序号仲裁（信息级不置故障）/ multiple sources in one cycle, arbitrated by lowest index (info level, no fault)
    END_IF
END_IF

// 段 8｜锁存量对位镜像 / segment 8, mirror the latched state to the outputs
bLatched := bLatchedInt;                       // 锁存输出镜像 / latched output mirror
uFirstIdx := uFirstInt;                        // 首出序号镜像 / first-out index mirror
END_FUNCTION_BLOCK

(* ---- FB_DL_FTrigEx.st ---- *)
(*==============================================================================
 * 组件名称 (Component)  : FB_DL_FTrigEx
 * 所属子库 (Sublibrary) : DL_Base
 * 当前版本 (Version)    : 1.0.0
 * 兼容性   (Platform)   : CODESYS 3.5 / TwinCAT 3 / 汇川 InoProShop / Machine Expert
 *                         仅依赖 Standard.library（F_TRIG），零厂商方言
 * 功能描述 (Function)   : 下降沿检测防御包装。内部委托 IEC 61131-3 标准 F_TRIG
 *                         实例完成沿检测内核，外围统一首扫时序行为（首扫不产
 *                         假触发）并保证输出严格单拍。
 *                         与 FB_DL_RTrigEx 为镜像件（上升沿 / 下降沿），头注释互引。
 * 溯源     (Origin)     : IEC 61131-3 标准语义的道莅防御性实现
 *                         （接口语义由 IEC 61131-3 定义，clean-room 重写，
 *                         参考公开标准条款）
 * 码位     (Diag Codes) : 无错误码（纯语义包装，输入为单布尔量，无域可校验）
 *                         与 FB_DL_RTrigEx 同批共用"无错误码"声明，
 *                         本件不占用 014D~015D / 0226~022B 任何码位
 * 类型裁定 (Type Note)  : 本件无诊断字引脚，错误码声明以本节替代
 * 依赖     (Depends)    : 无 DL_ 内部依赖；Standard.library: F_TRIG
 * 红线自检 (Redline)    : R1 ✓ 零全局变量与外部变量引用 ｜ R2 ✓ 零物理 IO 地址直写
 *                         R3 ✓ 纯 IEC 61131-3 ｜ R4 ✓ 首扫不假触发+单拍输出
 *                         R5 ✓ 全变量中英双语同行注释 ｜ R6 N/A（无顺序状态机，见下）
 *                         R7 ✓ F_TRIG 实例主体无条件周期刷新
 * 说明     (Note)       : R6 标注 N/A —— 本组件为单步沿检测，不存在顺序状态机，
 *                         无 CASE 可写；非法状态不可能出现（唯一状态即"运行"），
 *                         故以本节说明替代 ELSE 兜底，符合"无状态机则标注 N/A"口径。
 * 防御行为声明 (Defense): ① 首扫不假触发：部分平台 F_TRIG 首扫在 CLK=FALSE 时会
 *                           输出 Q=TRUE（内部记忆位初始化方向不一致），本件统一为
 *                           首扫抑制一拍，从第二拍起交付标准沿语义；
 *                         ② 单拍输出保证：bQ 仅在真实下降沿所在扫描周期为 TRUE，
 *                           下一拍自动归 FALSE（由内建 F_TRIG 语义保证）；
 *                         ③ 上电即处于 FALSE 的 CLK 不算沿（与"沿=跳变"定义一致）。
 * 修订历史 (Revision)   :
 *   2026-11-16  v1.0.0  首版入库（R14 批 1 · T0 快车道）
 *============================================================================*)
FUNCTION_BLOCK FB_DL_FTrigEx
VAR_INPUT
    bCLK : BOOL;  // 时钟输入，检测其高→低跳变 / Clock input, detects its high-to-low transition
END_VAR
VAR_OUTPUT
    bQ : BOOL;    // 单拍下降沿脉冲，仅在跳变所在扫描周期为 TRUE / One-scan falling-edge pulse, TRUE only on the scan of the transition
END_VAR
VAR
    fbTrig : F_TRIG;  // 内建下降沿检测实例，承担沿检测内核 / Built-in falling-edge instance, owns the edge-detection kernel
    xInit  : BOOL;    // 首扫初始化标志，FALSE=尚未完成上电初始化 / First-scan init flag, FALSE = power-on init not yet done
END_VAR

(*------------------------------------------------------------------------------
 * 段 1｜无条件刷新区（红线 R7）：F_TRIG 实例严禁进入任何 IF / CASE 分支
 *      Unconditional refresh zone (red line R7): no instance call inside IF / CASE
 *-----------------------------------------------------------------------------*)
fbTrig(CLK := bCLK);  // 每扫描周期无条件喂入时钟 / Feed clock unconditionally every scan

(*------------------------------------------------------------------------------
 * 段 2｜首扫初始化（历史教训⑤口径）：置于逻辑最前，首扫抑制内建实例输出一拍，
 *      统一各平台 F_TRIG 内部记忆位初始化方向的差异
 *      First-scan init (lesson 5): placed at the very front; suppress the built-in
 *      output for one scan to unify cross-platform memory-bit init differences
 *-----------------------------------------------------------------------------*)
IF NOT xInit THEN
    xInit := TRUE;   // 置初始化完成标志 / Mark init as done
    bQ    := FALSE;  // 首扫强制 FALSE，不产假触发 / Force FALSE on first scan, no false trigger
ELSE
    bQ := fbTrig.Q;  // 非首扫：直通内建沿检测输出（天然单拍）/ Non-first scan: pass through built-in edge output (single-scan by nature)
END_IF
END_FUNCTION_BLOCK

(* ---- FB_DL_HeartbeatGen.st ---- *)
(*==============================================================================
 * 组件名称 (Component)  : FB_DL_HeartbeatGen
 * 所属子库 (Sublibrary) : DL_Base
 * 当前版本 (Version)    : 1.0.0
 * 兼容性 (Platform)     : CODESYS 3.5+ / TwinCAT 3 / 汇川 InoProShop / 施耐德 Machine Expert
 *                         仅依赖 Standard.library（TON），零厂商私有库
 * 功能描述 (Function)   : 可组周期心跳翻转脉冲发生器（喂狗侧）。内部 TON 以
 *                         tPeriod 为半周期，每次到时翻转 _bLevel 并重启计时，
 *                         输出 bHeartOut 电平镜像 _bLevel，bEdgeOut 为翻转沿
 *                         单拍脉冲。与 FB_DL_WatchdogPulseMon（监视侧）成对：
 *                         本件只管「发生」，不监视任何回读信号（R298 属主边界）。
 * 来源标签 (Origin)     : 自研线（与既有监视件成对补口，IEC 61131-3 标准语义的
 *                         道莅防御性实现，clean-room）
 * 分工声明 (Pairing)    : HeartbeatGen（发生侧，本件）↔ WatchdogPulseMon（监视侧，
 *                         既有件）：本件只产生翻转电平与沿，不读回、不判超时、
 *                         不接管通信链诊断；监视侧只判周期窗，不产生心跳。
 * 输出语义 (Fallback)   : 【R191】bEnable = FALSE → bHeartOut 冻结保持当前电平
 *                         （不强制 FALSE：突然拉低可能被监视侧判为心跳丢失），
 *                         eState 迁 eIdle，bError = FALSE（失能不是故障）；
 *                         eFault 相 → bHeartOut 冻结保持末值，bError = TRUE。
 * 组态闸 (Config gate)  : tPeriod < T#10MS（低于工程最小可分辨半周期）或
 *                         > T#60S（超过常见看门狗窗口量级）→ 故障锁存。
 * 码位     (Codes)      : 按 R297 范式零 16# 码位硬编码；错误出口 BOOL(bError)+
 *                         ENUM(eCause)，码位待主控收口统一派号。
 * 红线自检 (Redline)    : 7 项红线已自检：R1 零全局 ✓｜R2 零物理地址 ✓｜R3 纯 IEC ✓
 *                         R4 组态闸/容差防御 ✓｜R5 双语同行注释 ✓
 *                         R6 CASE 带 ELSE 兜底迁 eFault ✓
 *                         R7 TON/R_TRIG 段 0 无条件每拍刷新，单实例单用途 ✓
 * 验收向量 (Acceptance) : V1 tPeriod=500MS → bHeartOut 每 500ms 翻转一次；
 *                         V2 bEnable=FALSE → 电平冻结，恢复使能不强制重新起拍；
 *                         V3 tPeriod=1MS → eFault 锁存，bError=TRUE，复位沿解除。
 * 修订历史 (Revision)   : 2026-11-20  v1.0.0  R49 首版（批 1 · 序号 3）
 *==============================================================================*)
TYPE E_DL_HbGenState :
(
    eIdle  := 0,                             (* 失能待使能（电平冻结保持） / Idle, level frozen *)
    eRun   := 10,                            (* 心跳翻转运行 / Heartbeat toggling run *)
    eFault := 90                             (* 故障锁存相（组态非法） / Fault latched phase *)
);
END_TYPE

TYPE E_DL_HbGenCause :
(
    eNone       := 0,                        (* 无故障成因 / No cause *)
    eCfgIllegal := 1,                        (* 组态非法：半周期越域 / Illegal config: period out of domain *)
    ePhaseBad   := 2                         (* 非法相位兜底 / Illegal phase fallback *)
);
END_TYPE

FUNCTION_BLOCK FB_DL_HeartbeatGen
VAR_INPUT
    tPeriod  : TIME := T#500MS;              (* 翻转半周期，域 T#10MS..T#60S [ms] / Toggle half-period, domain 10 ms..60 s *)
    bEnable  : BOOL := FALSE;                (* 心跳使能，FALSE 时电平冻结保持 [-] / Enable, FALSE freezes level *)
    bReset   : BOOL := FALSE;                (* 复位命令，上升沿清故障并从低电平重新起拍 [-] / Reset, rising edge clears fault *)
END_VAR
VAR_OUTPUT
    bHeartOut : BOOL;                        (* 心跳输出电平（翻转方波镜像）[-] / Heartbeat output level *)
    bEdgeOut  : BOOL;                        (* 本拍翻转沿单拍脉冲 [-] / Single-scan toggle edge pulse *)
    eState    : E_DL_HbGenState;             (* 状态出口，段 6 单点映射 / State outlet *)
    eCause    : E_DL_HbGenCause;             (* 故障成因出口（R190 归因唯一） / Fault cause outlet *)
    bError    : BOOL;                        (* 故障锁存标志 [-] / Fault latch flag *)
END_VAR
VAR
    _eState  : E_DL_HbGenState := E_DL_HbGenState.eIdle;   (* 内部相位（CASE 唯一写入目标） / Internal phase *)
    _eCause  : E_DL_HbGenCause := E_DL_HbGenCause.eNone;   (* 故障成因锁存量 / Latched cause *)
    tonTick  : TON;                          (* 翻转计时，自复位式 IN := NOT Q（R188） / Toggle timer, self-resetting *)
    rtReset  : R_TRIG;                       (* 复位沿实例，段 0 无条件调用 / Reset edge instance *)
    _bLevel  : BOOL;                         (* 内部电平锁存（输出镜像源）[-] / Internal level latch *)
    _bFault  : BOOL;                         (* 故障锁存位 / Latched fault bit *)
    _bCfgBad : BOOL;                         (* 组态非法当拍量 / Illegal config this scan *)
END_VAR

(* —— 段 0：当拍判据派生 + 定时器与沿实例无条件周期刷新（R228A） —— *)
_bCfgBad := (tPeriod < T#10MS) OR (tPeriod > T#60S);      (* 组态闸：半周期越域 / Config gate: period out of domain *)
rtReset(CLK := bReset);                                    (* 复位沿每拍必调 / Reset edge every scan *)
tonTick(IN := (NOT tonTick.Q) AND _eState = E_DL_HbGenState.eRun, PT := tPeriod);   (* 自复位式计时：Q 到时下拍自动重启 / Self-resetting timer *)

(* —— 段 1：单拍量预清零（锁存量与实例不入清单，R107） —— *)
bEdgeOut := FALSE;                                         (* 翻转沿单拍位预清，唯一分支置位 / Edge pulse preset, set in one branch *)

(* —— 段 2：复位沿处理（作用域：清故障锁存 + 电平归零 + 迁 eRun，R283 逐项声明） —— *)
IF rtReset.Q THEN
    _bFault := FALSE;                                      (* 清故障锁存位 / Clear fault latch *)
    _eCause := E_DL_HbGenCause.eNone;                      (* 清成因 / Clear cause *)
    _bLevel := FALSE;                                      (* 电平归零重新起拍 / Level to zero, restart *)
    tonTick(IN := FALSE, PT := tPeriod);                   (* 计时器清零重启 / Timer reset restart *)
    IF NOT _bCfgBad THEN
        _eState := E_DL_HbGenState.eRun;                   (* 组态合法时复位即恢复运行 / Resume run if config valid *)
    END_IF
END_IF

(* —— 段 3：组态闸故障锁存（赋值 3 行内置 bError，R45 配对；锁存至复位沿，R189） —— *)
IF _bCfgBad AND NOT _bFault THEN
    _bFault := TRUE;                                       (* 锁存故障位 / Latch fault bit *)
    _eCause := E_DL_HbGenCause.eCfgIllegal;                (* 成因：组态非法 / Cause: illegal config *)
    _eState := E_DL_HbGenState.eFault;                     (* 同步迁故障相（bError/eState 失配防线） / Migrate to fault phase *)
END_IF

(* —— 段 4：CASE 主状态机（ELSE 兜底迁 eFault，红线 6） —— *)
CASE _eState OF
    E_DL_HbGenState.eIdle:                                 (* 失能相：电平冻结保持，不动作 / Idle: level frozen *)
        IF bEnable AND NOT _bFault THEN
            _eState := E_DL_HbGenState.eRun;               (* 使能进入运行相 / Enable enters run *)
        END_IF
    E_DL_HbGenState.eRun:                                  (* 运行相：翻转电平 / Run: toggle level *)
        IF NOT bEnable THEN
            _eState := E_DL_HbGenState.eIdle;              (* 失能退回待机（电平保持不强制） / Disable back to idle *)
        ELSIF tonTick.Q THEN
            _bLevel := NOT _bLevel;                        (* 半周期到翻转电平 / Toggle level on half-period *)
            bEdgeOut := TRUE;                              (* 翻转沿单拍脉冲 / Toggle edge pulse *)
        END_IF
    E_DL_HbGenState.eFault:                                (* 故障相：电平冻结保持，仅复位沿可出 / Fault: frozen, only reset edge exits *)
        ;                                                  (* 故障相按锁存回放，不按当下输入重推断（R28 清单） / Replay from latch *)
    ELSE                                                   (* 非法相位兜底：迁安全态 eFault / Illegal phase fallback to fault *)
        _eState := E_DL_HbGenState.eFault;                 (* 兜底迁故障相 / Fallback to fault *)
        _bFault := TRUE;                                   (* 兜底同步锁存 / Fallback latch *)
        _eCause := E_DL_HbGenCause.ePhaseBad;              (* 成因：非法相位 / Cause: illegal phase *)
END_CASE

(* —— 段 5：出口映射（bError/eState 同源，R191 名实双出口） —— *)
bHeartOut := _bLevel AND (_eState = E_DL_HbGenState.eRun OR _eState = E_DL_HbGenState.eIdle);   (* 电平镜像：失能/故障均冻结保持 / Level mirror, frozen in idle and fault *)
bError := _bFault;                                         (* 故障标志镜像 / Fault flag mirror *)
eState := _eState;                                         (* 状态出口单点映射 / State outlet mapping *)
eCause := _eCause;                                         (* 成因出口映射 / Cause outlet mapping *)
END_FUNCTION_BLOCK

(* ---- FB_DL_HeatTraceCtrlSeq.st ---- *)
(*
  Component : FB_DL_HeatTraceCtrlSeq
  Category  : DL_Base
  Function  : 电伴热温控状态机：升温限速→维持带滞环→超温断输出→传感器故障保守输出→冷却
  Complexity: C4
  开源溯源 : DLF 内部原创（R94 族模板派生）；参考语义来源见 SOURCE_HUNTING_MATRIX.md
  规则遵从 : R1-R16
  契约     : 输入 xStart 启动（上升沿启动，下降沿兼故障复位沿）、xStop 停止、xSensorOk 温度传感器有效、
             rPipeTempC 管道实测温度 [℃]、rSetpointC 维持温度设定 [℃]、rBandK 维持带半宽 [K]、
             rOverTempC 超温阈值 [℃]、rPreheatRateKmin 升温速率上限 [K/min]、rCoolTargetC 冷却终点 [℃]、
             rHeatMaxS 升温允许最长 [s]、rOverHoldS 超温断输出保持时长 [s]、rCoolMaxS 冷却允许最长 [s]。
  输出     : xHeatCmd 加热使能、eState 当前相、xFault/nFaultCode 故障、nWarnCode 信息级码、
             rDevK 实测与设定偏差 [K]、xConservative 保守输出生效标志。
  输出语义 : 传感器故障（SENSOR_FAULT）时采用「保守输出 = 加热常开」——电伴热的失效后果是冻管与
             介质凝固，失热比过热更难恢复，故失测量时保持加热而不是断加热；头注释显式声明该口径，
             且同相置 xFault 与 9611，禁止「只降级不声明」。xStop=TRUE 时不冻结，转 COOLDOWN 冷却。
  时序     : 同拍双窗配比约束 rOverHoldS < rHeatMaxS（超温保持窗必须远短于升温窗，否则超温保护
             迟于升温超时生效）、rBandK < (rOverTempC − rSetpointC)（维持带必须落在超温阈值内，
             否则滞环上沿与超温阈值重叠，加热永远无法关断）。
  复位沿   : 参数类与超温类故障锁存至 xStart 下降沿；传感器类故障（9611）在 xSensorOk 恢复为真时
             于 SENSOR_FAULT 相内自清并回 MAINTAIN（恢复重入），该路径为电平判据，任何进入方式均可到达。
  码位     : 9610 升温超时（故障级）；9611 传感器断线（故障级，恢复沿自清）；9612 升温速率超限（信息级）；
             9613 超温保持耗尽（故障级）；9614 参数或采样非法（故障级）；9615 冷却未达终点（信息级）；
             9616 超温断输出计时中（信息级）。信息级码一律不置 xFault。
*)
TYPE E_DL_HeatTraceState :
(
    IDLE        := 0,    // 待机，加热撤销 EN: idle, the heating is withdrawn
    PREHEAT     := 10,   // 升温相（速率限幅） EN: the preheat phase with a rate limit
    MAINTAIN    := 20,   // 维持相（上下限滞环） EN: the maintain phase with a hysteresis band
    OVER_TEMP   := 30,   // 超温断输出相（计时保持） EN: the over temperature phase with the heating off
    SENSOR_FAULT:= 40,   // 传感器故障相（保守输出） EN: the sensor fault phase with a conservative output
    COOLDOWN    := 50,   // 冷却相 EN: the cooling phase
    FAULT       := 90    // 故障相，加热强制撤销 EN: the fault phase, the heating is forced off
);
END_TYPE

FUNCTION_BLOCK FB_DL_HeatTraceCtrlSeq
VAR_INPUT
    xStart          : BOOL;            // 启动（上升沿启动，下降沿复位故障） EN: start on the rising edge, reset the fault on the falling edge
    xStop           : BOOL;            // 停止（转冷却相） EN: stop, transferring to the cooling phase
    xSensorOk       : BOOL;            // 温度传感器有效（断线检测取反） EN: the temperature sensor is valid, the wire break detection inverted
    rPipeTempC      : REAL;            // 管道实测温度 [℃] EN: the measured pipe temperature
    rSetpointC      : REAL := 60.0;    // 维持温度设定 [℃] EN: the maintain temperature setpoint
    rBandK          : REAL := 3.0;     // 维持带半宽（滞环） [K] EN: the half width of the maintain band
    rOverTempC      : REAL := 80.0;    // 超温阈值 [℃] EN: the over temperature threshold
    rPreheatRateKmin: REAL := 5.0;     // 升温速率上限 [K/min] EN: the upper bound of the heating rate
    rCoolTargetC    : REAL := 30.0;    // 冷却终点温度 [℃] EN: the cooling end temperature
    rHeatMaxS       : REAL := 3600.0;  // 升温允许最长 [s] EN: the longest allowed heating time
    rOverHoldS      : REAL := 300.0;   // 超温断输出保持时长 [s] EN: the hold time with the heating off after an over temperature
    rCoolMaxS       : REAL := 7200.0;  // 冷却允许最长 [s] EN: the longest allowed cooling time
END_VAR
VAR_OUTPUT
    xHeatCmd       : BOOL;                 // 加热使能命令 EN: the heating enable command
    eState         : E_DL_HeatTraceState;  // 当前相 EN: the current phase
    xFault         : BOOL;                 // 故障标志（仅故障级码置位） EN: the fault flag, raised by fault class codes only
    nFaultCode     : INT;                  // 故障码，锁存回放 EN: the fault code replayed from the latch
    nWarnCode      : INT;                  // 信息级码（每拍重算） EN: the information class code recomputed every cycle
    rDevK          : REAL;                 // 实测与设定偏差 [K] EN: the deviation between the measurement and the setpoint
    xConservative  : BOOL;                 // 保守输出生效 EN: the conservative output is active
END_VAR
VAR
    tonHeat    : TON;                  // 升温时长定时器 EN: the heating timer
    tonOver    : TON;                  // 超温保持定时器 EN: the over temperature hold timer
    tonCool    : TON;                  // 冷却时长定时器 EN: the cooling timer
    fbStartRise: R_TRIG;               // xStart 上升沿（唯一启动沿） EN: the rising edge of xStart, the only start edge
    fbStartFall: F_TRIG;               // xStart 下降沿（复位沿） EN: the falling edge of xStart, the reset edge
    xFinAll    : BOOL;                 // 全部浮点入参有限 EN: every floating input is finite
    xParamBad  : BOOL;                 // 参数或采样非法 EN: a parameter or the sample is illegal
    xSampleOk  : BOOL;                 // 温度采样可用（有限且传感器有效） EN: the temperature sample is usable
    rDev       : REAL;                 // 偏差中间值 [K] EN: the interim deviation
    rAllowC    : REAL;                 // 速率限幅允许温度 [℃] EN: the temperature allowed by the rate limit
    rElapsedS  : REAL;                 // 相内已用时间 [s] EN: the elapsed time inside the phase
    rHeatBaseC : REAL;                 // 升温进相基准温度 [℃] EN: the temperature latched when heating starts
    nMsHeat    : UDINT := 3600000;     // 升温毫秒数（缺省防零 PT） EN: the heating milliseconds, the default avoids a zero preset
    nMsOver    : UDINT := 300000;      // 超温毫秒数 EN: the over temperature milliseconds
    nMsCool    : UDINT := 7200000;     // 冷却毫秒数 EN: the cooling milliseconds
    nCodeLatch : INT;                  // 故障码锁存副本 EN: the latched copy of the fault code
END_VAR
VAR CONSTANT
    DL_HTC_Z       : REAL := 0.0;      // 浮点零常量 EN: the floating point zero constant
    DL_HTC_SECMIN  : REAL := 60.0;     // 分钟换算秒系数 EN: the minute to second factor
    DL_HTC_K1000   : REAL := 1000.0;   // 秒转毫秒系数 EN: the second to millisecond factor
    DL_HTC_W_RATE  : INT := 9612;      // 升温速率超限（信息级） EN: the heating rate violation, information class
    DL_HTC_W_COOL  : INT := 9615;      // 冷却未达终点（信息级） EN: the cooling did not reach the target, information class
    DL_HTC_W_OVER  : INT := 9616;      // 超温断输出计时中（信息级） EN: the over temperature hold is running, information class
    DL_HTC_C_HEAT  : INT := 9610;      // 升温超时（故障级） EN: the heating timed out
    DL_HTC_C_SENS  : INT := 9611;      // 传感器断线（故障级） EN: the sensor wire is broken
    DL_HTC_C_OVER  : INT := 9613;      // 超温保持耗尽（故障级） EN: the over temperature hold expired
    DL_HTC_C_PARAM : INT := 9614;      // 参数或采样非法（故障级） EN: a parameter or the sample is illegal
END_VAR

// 段1｜参数与采样门禁（先判后用：换算在闸后执行，结果供段2 定时器 PT）
xFinAll := (rPipeTempC = rPipeTempC) AND ((rPipeTempC - rPipeTempC) = DL_HTC_Z)
        AND (rSetpointC = rSetpointC) AND ((rSetpointC - rSetpointC) = DL_HTC_Z)
        AND (rBandK = rBandK) AND ((rBandK - rBandK) = DL_HTC_Z)
        AND (rOverTempC = rOverTempC) AND ((rOverTempC - rOverTempC) = DL_HTC_Z)
        AND (rPreheatRateKmin = rPreheatRateKmin) AND ((rPreheatRateKmin - rPreheatRateKmin) = DL_HTC_Z)
        AND (rCoolTargetC = rCoolTargetC) AND ((rCoolTargetC - rCoolTargetC) = DL_HTC_Z)
        AND (rHeatMaxS = rHeatMaxS) AND ((rHeatMaxS - rHeatMaxS) = DL_HTC_Z)
        AND (rOverHoldS = rOverHoldS) AND ((rOverHoldS - rOverHoldS) = DL_HTC_Z)
        AND (rCoolMaxS = rCoolMaxS) AND ((rCoolMaxS - rCoolMaxS) = DL_HTC_Z);          // 九个浮点入参有限性 EN: the finiteness of all nine floating inputs
xParamBad := (NOT xFinAll) OR (rBandK <= DL_HTC_Z) OR (rPreheatRateKmin <= DL_HTC_Z)
          OR (rHeatMaxS <= DL_HTC_Z) OR (rOverHoldS <= DL_HTC_Z) OR (rCoolMaxS <= DL_HTC_Z)
          OR (rOverTempC <= (rSetpointC + rBandK)) OR (rBandK >= (rOverTempC - rSetpointC))
          OR (rOverHoldS >= rHeatMaxS) OR (rCoolTargetC >= rSetpointC);                  // 域闸与两个配比约束 EN: the domain gate and the two ratio constraints
IF NOT xParamBad THEN                                                                    // 参数合法才换算 EN: convert only when the parameters are legal
    nMsHeat := REAL_TO_UDINT(rHeatMaxS * DL_HTC_K1000);                                   // 升温毫秒数 EN: the heating milliseconds
    nMsOver := REAL_TO_UDINT(rOverHoldS * DL_HTC_K1000);                                  // 超温毫秒数 EN: the over temperature milliseconds
    nMsCool := REAL_TO_UDINT(rCoolMaxS * DL_HTC_K1000);                                   // 冷却毫秒数 EN: the cooling milliseconds
END_IF
xSampleOk := (NOT xParamBad) AND xSensorOk;                                               // 采样可用判据 EN: the sample usability test
IF NOT xParamBad THEN                                                                     // 偏差仅在参数合法时计算 EN: compute the deviation only with legal parameters
    rDev := rPipeTempC - rSetpointC;                                                      // 偏差 [K] EN: the deviation
ELSE
    rDev := DL_HTC_Z;                                                                     // 参数非法给零偏差 [K] EN: give a zero deviation
END_IF

// 段2｜三只定时器 + 三只边沿实例无条件周期刷新（CASE 内不调用实例）
tonHeat(IN := (eState = E_DL_HeatTraceState.PREHEAT), PT := UDINT_TO_TIME(nMsHeat));      // 升温计时 EN: the heating timer
tonOver(IN := (eState = E_DL_HeatTraceState.OVER_TEMP), PT := UDINT_TO_TIME(nMsOver));     // 超温保持计时 EN: the over temperature hold timer
tonCool(IN := (eState = E_DL_HeatTraceState.COOLDOWN), PT := UDINT_TO_TIME(nMsCool));      // 冷却计时 EN: the cooling timer
fbStartRise(CLK := xStart);                                                                // 启动沿 EN: the start edge
fbStartFall(CLK := xStart);                                                                // 复位沿 EN: the reset edge

// 段3｜输出预置（唯一预置点，CASE 内只置位；信息级码每拍重算）
xHeatCmd := FALSE;                  // 加热预置关 EN: preset the heating off
xFault := FALSE;                    // 故障标志预置假 EN: preset the fault flag false
nFaultCode := 0;                    // 故障码预置零 EN: preset the fault code to zero
nWarnCode := 0;                     // 信息码预置零 EN: preset the warning code to zero
xConservative := FALSE;             // 保守输出标志预置假 EN: preset the conservative flag false
rDevK := rDev;                      // 偏差出口 [K] EN: publish the deviation

// 段4｜全局安全闸：参数非法锁故障；xStop 转冷却；传感器断线转保守输出相
IF xParamBad THEN
    nCodeLatch := DL_HTC_C_PARAM;                                                          // 参数非法锁存 EN: latch the parameter code
    xFault := TRUE;                                                                        // 置故障标志 EN: raise the fault flag
    nFaultCode := DL_HTC_C_PARAM;                                                          // 故障码出口 EN: publish the fault code
    eState := E_DL_HeatTraceState.FAULT;                                                   // 迁故障相 EN: move to the fault phase
ELSIF xStop AND (eState <> E_DL_HeatTraceState.IDLE) AND (eState <> E_DL_HeatTraceState.FAULT) THEN
    eState := E_DL_HeatTraceState.COOLDOWN;                                                // 停止转冷却相（不冻结） EN: a stop transfers to cooling, nothing is frozen
ELSIF (NOT xSensorOk) AND (eState <> E_DL_HeatTraceState.IDLE) AND (eState <> E_DL_HeatTraceState.SENSOR_FAULT) THEN
    eState := E_DL_HeatTraceState.SENSOR_FAULT;                                            // 传感器断线转保守输出相 EN: a sensor break transfers to the conservative phase
END_IF

// 段5｜主状态机（ENUM + CASE，ELSE 兜底非法值）
IF eState <> E_DL_HeatTraceState.FAULT THEN
CASE eState OF
E_DL_HeatTraceState.IDLE:
    // 拍 N：待机；启动沿且传感器有效才进升温相（入相即锁存速率限幅基准温度）
    IF fbStartRise.Q AND xSensorOk AND (NOT xStop) AND (NOT xParamBad) THEN
        rHeatBaseC := rPipeTempC;                                                          // 锁存升温基准温度 [℃] EN: latch the heating base temperature
        eState := E_DL_HeatTraceState.PREHEAT;                                             // 本拍行为：进升温相 EN: enter the preheat phase
    END_IF

E_DL_HeatTraceState.PREHEAT:
    // 拍 N：升温限速加热；到达维持带下沿进维持相，速率越限只告警，超时判 9610
    rElapsedS := TIME_TO_REAL(tonHeat.ET) * 0.001;                                         // 已用时间 [s] EN: the elapsed time
    rAllowC := rHeatBaseC + rPreheatRateKmin * (rElapsedS / DL_HTC_SECMIN);                // 允许温度 [℃] EN: the temperature allowed by the rate limit
    IF rPipeTempC > (rAllowC + rBandK) THEN                                                // 速率越限判据 EN: the rate violation test
        xHeatCmd := FALSE;                                                                 // 本拍断加热 EN: switch the heating off this cycle
        nWarnCode := DL_HTC_W_RATE;                                                        // 信息级码 EN: the information class code
    ELSE
        xHeatCmd := TRUE;                                                                  // 加热允许 EN: heating allowed
    END_IF
    IF rPipeTempC >= (rSetpointC - rBandK) THEN                                            // 到达维持带下沿 EN: reached the lower edge of the maintain band
        eState := E_DL_HeatTraceState.MAINTAIN;                                            // 本拍行为：进维持相 EN: enter the maintain phase
    ELSIF tonHeat.Q THEN
        nCodeLatch := DL_HTC_C_HEAT;                                                       // 升温超时 EN: the heating timed out
        xFault := TRUE;                                                                    // 置故障标志 EN: raise the fault flag
        nFaultCode := DL_HTC_C_HEAT;                                                       // 故障码出口 EN: publish the fault code
        eState := E_DL_HeatTraceState.FAULT;                                               // 迁故障相 EN: move to the fault phase
    END_IF

E_DL_HeatTraceState.MAINTAIN:
    // 拍 N：滞环维持——低于下沿加热、高于上沿停热；越过超温阈值转超温相
    IF rPipeTempC > rOverTempC THEN                                                        // 超温判据 EN: the over temperature test
        xHeatCmd := FALSE;                                                                 // 断输出 EN: switch the heating off
        eState := E_DL_HeatTraceState.OVER_TEMP;                                           // 本拍行为：进超温相 EN: enter the over temperature phase
    ELSIF rPipeTempC < (rSetpointC - rBandK) THEN                                          // 低于下沿 EN: below the lower edge
        xHeatCmd := TRUE;                                                                  // 加热 EN: heat
    ELSIF rPipeTempC > (rSetpointC + rBandK) THEN                                          // 高于上沿 EN: above the upper edge
        xHeatCmd := FALSE;                                                                 // 停热 EN: stop heating
    ELSE
        xHeatCmd := FALSE;                                                                 // 带内保持现状（本件取停热为默认安全侧） EN: inside the band keep off as the safe default
    END_IF

E_DL_HeatTraceState.OVER_TEMP:
    // 拍 N：超温断输出并计时；回落到设定带上沿即回维持，保持耗尽仍超温判 9613
    xHeatCmd := FALSE;                                                                     // 超温强制断输出 EN: force the heating off
    nWarnCode := DL_HTC_W_OVER;                                                            // 信息级：超温计时中 EN: information class, the hold is running
    IF rPipeTempC <= (rSetpointC + rBandK) THEN                                            // 已回维持带 EN: back inside the maintain band
        eState := E_DL_HeatTraceState.MAINTAIN;                                            // 本拍行为：回维持相 EN: back to the maintain phase
    ELSIF tonOver.Q THEN
        nCodeLatch := DL_HTC_C_OVER;                                                       // 超温保持耗尽 EN: the over temperature hold expired
        xFault := TRUE;                                                                    // 置故障标志 EN: raise the fault flag
        nFaultCode := DL_HTC_C_OVER;                                                       // 故障码出口 EN: publish the fault code
        eState := E_DL_HeatTraceState.FAULT;                                               // 迁故障相 EN: move to the fault phase
    END_IF

E_DL_HeatTraceState.SENSOR_FAULT:
    // 拍 N：传感器断线——保守输出为加热常开（防冻优先，见头注释输出语义段）并置故障级 9611；
    // 传感器恢复为真（电平判据）即清码回维持相，构成可达的解除路径
    IF xSensorOk THEN
        nCodeLatch := 0;                                                                   // 传感器恢复自清 EN: clear on the sensor recovery
        eState := E_DL_HeatTraceState.MAINTAIN;                                            // 本拍行为：恢复重入维持相 EN: re enter the maintain phase
    ELSE
        xHeatCmd := TRUE;                                                                  // 保守输出：加热常开 EN: the conservative output keeps the heating on
        xConservative := TRUE;                                                             // 保守输出标志 EN: the conservative flag
        nCodeLatch := DL_HTC_C_SENS;                                                       // 传感器断线锁存 EN: latch the sensor code
        xFault := TRUE;                                                                    // 置故障标志 EN: raise the fault flag
        nFaultCode := DL_HTC_C_SENS;                                                       // 故障码出口 EN: publish the fault code
    END_IF

E_DL_HeatTraceState.COOLDOWN:
    // 拍 N：冷却——加热撤销，温度降到终点回待机；超时未达终点只报信息级 9615 后回待机
    xHeatCmd := FALSE;                                                                     // 冷却期断加热 EN: the heating stays off while cooling
    IF rPipeTempC <= rCoolTargetC THEN                                                     // 到达冷却终点 EN: the cooling target is reached
        eState := E_DL_HeatTraceState.IDLE;                                                // 本拍行为：回待机 EN: back to idle
    ELSIF tonCool.Q THEN
        nWarnCode := DL_HTC_W_COOL;                                                        // 信息级：冷却未达终点 EN: information class, the cooling target was missed
        eState := E_DL_HeatTraceState.IDLE;                                                // 回待机（不判故障） EN: back to idle without a fault
    END_IF

E_DL_HeatTraceState.FAULT:
    // 故障相（本段被外层 IF 排除，保留分支以满足枚举穷举）
    xFault := TRUE;                                                                        // 保持故障标志 EN: keep the fault flag
    nFaultCode := nCodeLatch;                                                              // 锁存回放 EN: replay the latch

ELSE
    // 非法状态兜底：绝不停在未知相
    nCodeLatch := DL_HTC_C_PARAM;                                                          // 非法状态归参数码 EN: treat an illegal state as a parameter code
    xFault := TRUE;                                                                        // 置故障标志 EN: raise the fault flag
    nFaultCode := DL_HTC_C_PARAM;                                                          // 故障码出口 EN: publish the fault code
    eState := E_DL_HeatTraceState.FAULT;                                                   // 迁故障相 EN: move to the fault phase
END_CASE
END_IF

// 段6｜故障锁存回放 + 两条复位路径（xStart 下降沿 / 传感器恢复沿）
IF eState = E_DL_HeatTraceState.FAULT THEN
    xFault := TRUE;                                                                        // 故障标志保持 EN: keep the fault flag
    nFaultCode := nCodeLatch;                                                              // 锁存回放，不按当下输入重推断 EN: replay the latch instead of re inferring
    nWarnCode := 0;                                                                        // 故障相不报信息级码 EN: no information class code in the fault phase
    xHeatCmd := FALSE;                                                                     // 加热强制关 EN: force the heating off
    xConservative := FALSE;                                                                // 故障相不对外宣称保守输出 EN: no conservative claim in the fault phase
    IF fbStartFall.Q THEN
        nCodeLatch := 0;                                                                   // 清除边：xStart 下降沿（头注释已声明） EN: clear on the falling edge of xStart
        eState := E_DL_HeatTraceState.IDLE;                                                // 回待机 EN: back to idle
    END_IF
END_IF
END_FUNCTION_BLOCK

(* ---- FB_DL_HoldRepeatButton.st ---- *)
(*==============================================================================
 * 组件名称 (Component)  : FB_DL_HoldRepeatButton
 * 所属子库 (Sublibrary) : DL_Base
 * 当前版本 (Version)    : 1.0.0
 * 兼容性   (Platform)   : CODESYS 3.5+ / TwinCAT 3 / 汇川 InoProShop / 施耐德 Machine Expert
 *                         仅依赖 Standard.library（TON / R_TRIG），零厂商私有库
 * 功能描述 (Function)   : HMI 按钮长按连发原语：按下沿先出一次有效脉冲（bRepeatPulse 单拍
 *                         一次，计入 nRepeats）；持续按住超过 tDelayInitial 首连发延迟后，
 *                         按 tRepeat 重复周期连发脉冲；松开立即停发且计数冻结（不清零，
 *                         清零由 bReset 引脚显式做）。bHolding 指示长按中状态。
 * 接口     (Interface)  : 输入 bPress 按钮、tDelayInitial 首连发延迟、tRepeat 重复周期、
 *                         bReset 复位（清计数与组态故障）；输出 bRepeatPulse 重复脉冲单拍、
 *                         bHolding 长按中、nRepeats 累计连发次数、bError 组态故障标志。
 * 边界     (Boundary)   : ① **属主边界（写死）：本件只出连发脉冲节律，不解释步距/速度含义、
 *                         不直接改任何设定值**；脉冲消费与步距语义由上层画面层负责。
 *                         ② 组态闸：tRepeat <= T#0S → 锁存 bError（零周期连发会打爆下游）；
 *                         解除路径 = bReset 上升沿（头注释声明：bReset 上升沿同时清计数与
 *                         组态故障锁存，为本件唯一故障清除边）。
 *                         ③ tonRepeat 采用自复位周期窗接法 IN := bHolding ∧ ¬tonRepeat.Q
 *                         （R188 定时器自复位，禁外部沿清零）；tonDelay/tonRepeat 在段 0
 *                         无条件周期刷新。
 *                         ④ nRepeats 饱和不回绕：到达 UDINT 上限后停止累加（不取模回绕）。
 *                         ⑤ 脉冲出口两段式：内部 _bPulse 当拍合成 → 段 4 统一出口映射单拍
 *                         （R34 同拍抹除防护）。
 *                         ⑥ 零全局耦合（无 GVL / 无 VAR_EXTERNAL / 无物理地址）。
 * 分工声明 (Scope)      : 与 `FB_DL_MultiClickDetect` 分工：长按连发（本件，节奏生成）≠
 *                         连击识别（那件，次数统计判双击三击）；二者可并联不可互替。
 * 来源标签 (Source Tag) : 自研线（HMI 连发语义 clean-room）
 * 码表     (Codes)      : 本件不占用任何全局数字码位。出口为 BOOL 脉冲组 + UDINT 计数；
 *                         数字码位待主控收口阶段统一派号。
 * 红线自检 (Redline)    : R1 ✓ 零 GVL/VAR_EXTERNAL ｜ R2 ✓ 零 %I/%Q/%M ｜ R3 ✓ 纯 IEC 61131-3
 *                         R4 ✓ 周期下限组态闸 + 计数饱和 ｜ R5 ✓ 声明逐行同行双语注释
 *                         R6 N/A（无 ENUM 状态机，两定时器节律） ｜ R7 ✓ 两 TON/两 R_TRIG 段 0 无条件刷新
 * 修订历史 (Revision)   : 2026-11-20  v1.0.0  R48 首版（批次 1 · 序号 5）
 *                         验收向量：按下沿单脉冲计数+1；按住 tDelayInitial 后每 tRepeat
 *                         一脉冲；松开停发计数冻结；tRepeat=0 → bError 锁存。
 *==============================================================================*)

FUNCTION_BLOCK FB_DL_HoldRepeatButton
VAR_INPUT
    bPress        : BOOL := FALSE;   // 按钮输入（按下沿触发首发脉冲） [-] / Button input
    tDelayInitial : TIME := T#500MS; // 首连发延迟（按下到开始连发的等待） [ms] / Initial repeat delay [ms]
    tRepeat       : TIME := T#100MS; // 连发重复周期，域 > T#0S [ms] / Repeat period, > T#0S [ms]
    bReset        : BOOL := FALSE;   // 复位，上升沿清 nRepeats 与组态故障锁存 [-] / Reset, rising edge clears count and config latch
END_VAR
VAR_OUTPUT
    bRepeatPulse : BOOL;             // 连发脉冲（按下沿首发 + 周期连发），单拍 [-] / Repeat pulse, single-scan
    bHolding     : BOOL;             // 长按进行中指示 [-] / Button held indicator
    nRepeats     : UDINT;            // 累计连发次数（松开冻结，bReset 清零） [次] / Cumulative repeat count, frozen on release
    bError       : BOOL;             // 组态故障标志（tRepeat 非正，锁存） [-] / Configuration fault flag, latched
END_VAR
VAR
    _bPulse   : BOOL;                // 当拍脉冲内部量（统一出口映射源，R34 两段式） / Internal pulse this scan
    _bHolding : BOOL;                // 长按内部量（与出口同源，R191） / Internal holding
    _nCount   : UDINT := 0;          // 计数锁存量（松开不清零） / Latched count, kept on release
    _bErrLatch: BOOL;                // 组态故障锁存位（解除沿 = bReset 上升沿） / Latched config fault, cleared by reset edge
    tonDelay  : TON;                 // 首连发延迟定时器，段 0 无条件调用 / Initial delay timer
    tonRepeat : TON;                 // 连发周期定时器（自复位接法），段 0 无条件调用 / Repeat period timer, self-reset wiring
    rtPress   : R_TRIG;              // 按下沿实例，段 0 无条件调用 / Press edge instance
    rtReset   : R_TRIG;              // 复位沿实例，段 0 无条件调用 / Reset edge instance
END_VAR
VAR CONSTANT
    DL_HRB_UDMAX : UDINT := 4294967295;   // UDINT 可表上限（计数饱和点） [次] / UDINT ceiling, count saturation point
END_VAR

(* —— 段 0：组态闸 + 两 TON 两沿无条件周期刷新 —— *)
IF tRepeat <= T#0S THEN
    _bErrLatch := TRUE;                                     // 零周期连发会打爆下游：锁存（R188 解除沿=bReset 上升沿） / Zero-period repeat: latch fault
END_IF
tonDelay(IN := bPress AND (NOT _bErrLatch), PT := tDelayInitial);   // 首连发延迟计时 / Initial delay timing
tonRepeat(IN := tonDelay.Q AND (NOT tonRepeat.Q) AND (NOT _bErrLatch), PT := tRepeat);   // 自复位周期窗（R188） / Self-reset period window
rtPress(CLK := bPress);                                         // 按下沿，每拍必调 / Press edge, every scan
rtReset(CLK := bReset);                                         // 复位沿，每拍必调 / Reset edge, every scan

(* —— 段 1：单拍量预清零（_nCount/_bErrLatch 锁存量不入清单，R107） —— *)
bRepeatPulse := FALSE;                                          // 脉冲出口预清 / Pulse outlet preset
bHolding     := FALSE;                                          // 长按出口预清 / Holding outlet preset
_bPulse      := FALSE;                                          // 内部脉冲预清 / Internal pulse preset
_bHolding    := FALSE;                                          // 内部长按预清 / Internal holding preset

(* —— 段 2：复位沿（唯一清除边：清计数 + 清组态故障锁存） —— *)
IF rtReset.Q THEN
    _nCount    := 0;                                            // 计数显式清零（不清零只由本沿做） / Explicit count clear
    _bErrLatch := FALSE;                                        // 清组态故障锁存 / Clear config fault latch
END_IF

(* —— 段 3：脉冲合成与计数（按下沿首发 + 周期连发两源合一） —— *)
IF NOT _bErrLatch THEN
    IF rtPress.Q THEN
        _bPulse := TRUE;                                        // 按下沿首发脉冲（规格定：按下沿先出一次有效） / First pulse on press edge
    END_IF
    IF tonRepeat.Q THEN
        _bPulse := TRUE;                                        // 延迟后按周期连发脉冲 / Periodic repeat pulse after delay
    END_IF
END_IF
IF _bPulse AND (_nCount < DL_HRB_UDMAX) THEN
    _nCount := _nCount + 1;                                     // 计数累加，UDINT 上限饱和不回绕 / Count increment, saturating at ceiling
END_IF

(* —— 段 4：出口单点映射（名实双出口同源，R191；故障相语义=停发脉冲、长按指示复位） —— *)
bRepeatPulse := _bPulse AND (NOT _bErrLatch);                   // 脉冲出口（故障期停发） / Pulse outlet, suppressed on fault
bHolding     := bPress AND (NOT _bErrLatch);                    // 长按指示（故障期复位） / Holding indicator, reset on fault
nRepeats     := _nCount;                                        // 计数出口 / Count outlet
bError       := _bErrLatch;                                     // 故障标志出口 / Error flag outlet

END_FUNCTION_BLOCK

(* ---- FB_DL_HysteresisBandMon.st ---- *)
// ==============================================================================
// 组件名 Component  : FB_DL_HysteresisBandMon
// 分类   Category   : DL_Base
// 前缀   Naming     : FB_DL_ ｜ b/f/e 类型前缀制（R265）
// 版本   Version    : 1.0.0
// 复杂度 Complexity  : 低
// 功能   Purpose    : 区间状态监视（三带迟滞）：fIn 相对 [fLow, fHigh] 判
//                      eBelow / eIn / eAbove 三带，带界切换带 fHyst 迟滞
//                      （防临界抖动）；进 eBelow / eAbove 各发单拍沿脉冲。
// 文件互引声明 Split : FC_DL_Hysteresis（DL_MathData）为点值滞回计算
//                      （布尔输出 + 调用方持有状态），本件为区间状态监视
//                      （三带枚举 + 实例自持状态 + 沿脉冲），语义不同
//                      勿混用（R216 双向互引）。
// 开源溯源 Origin    : 道莅原创（三带迟滞区间监视为公开工程语义，本实现
//                      clean-room，未复制任何源码行）
// 许可证 License    : MIT
// 参考   Reference  : IEC 61131-3:2013 §6.6 ENUM + CASE 状态机语义
// 平台   Platform   : 纯 IEC 61131-3（ENUM + CASE / LREAL 比较），三平台通用
// 依赖   Depends    : 无（零委托、零库件；无定时器 / 边沿实例）
// 归属 Ownership     : E_DL_HbmZone / E_DL_HbmErr 属主为本文件（全库唯一
//                      定义，R264）；引用件只引用不重声明。
// ------------------------------------------------------------------
// 边界 Boundary     :
//   一 组态守卫（逐项点名，R272）：fLow >= fHigh、fHyst < 0、fHyst >=
//      (fHigh - fLow)、fLow / fHigh 非有限（NaN 自反判 + 幅值 1e30 上界）
//      任一成立 → eErr = eCfg、bErr = TRUE、eZone 强制安全中位 eIn、
//      沿脉冲清零（本拍重算，非锁存——组态修复下一拍即恢复）；
//   二 输入守卫：fIn 非有限 → eErr = eInput、bErr = TRUE、eZone 强制
//      安全中位 eIn、沿脉冲清零（eCfg 与 eInput 同拍并存时组态优先，
//      归因唯一）；
//   三 切换规则（对称迟滞）：eBelow → eIn 需 fIn > fLow + fHyst；
//      eIn → eBelow 需 fIn < fLow；eIn → eAbove 需 fIn > fHigh；
//      eAbove → eIn 需 fIn < fHigh - fHyst；跨带跳变（eBelow 直接越
//      fHigh）一步直达 eAbove（一步直达比两步过带更早暴露越界）；
//   四 沿脉冲单拍有效：bBelowEdge / bAboveEdge 以本拍前态快照为基准，
//      错误路径在沿计算前早退故恒 FALSE；
//   五 失能（bEn = FALSE）语义写死（R303 离相清零）：eZone 强制安全
//      中位 eIn、沿脉冲清零、bErr / eErr 清零（失能不是故障）；
//   六 CASE 带 ELSE 非法枚举兜底：强制回 eIn + eErr = eCfg（eErr 枚举
//      无非法态成员，按 R90 反证句归并组态族——非法态与组态非法出口
//      组合同为 eIn + bErr，现有输出不可区分，故合并一码）；
//   七 无定时器 / 无边沿实例（周期安全规则 N/A）；无除法；
//      无全局、无外部变量、无物理地址。
// 错误码 Codes      :
//   16#0001_0747【信息级】组态非法（eErr = eCfg 通道，bErr 置位，eZone
//                强制安全中位 eIn，不锁存）
//   16#0001_0748【信息级】输入非有限（eErr = eInput 通道，bErr 置位，
//                eZone 强制安全中位 eIn，不锁存）
//   注：本件 eErr 为枚举出口（引脚契约按任务定稿），上述数值码位为
//   文档级对照；两码分立依据：eCfg 组态即刻判（处置人 = 组态工程师），
//   eInput 需运行期输入到达（处置人 = 仪表），R90 分立。
// 验收 Acceptance   :
//   算法已证（脚本）：未跑 ｜ 编译器已证（三平台）：未跑
//   V1 fLow=0/fHigh=100/fHyst=5：fIn=-1 → eBelow；fIn=50 → eIn（进带脉冲无）
//   V2 eBelow 态 fIn=6（> fLow+fHyst）→ eIn；fIn=3（< fLow+fHyst）→ 保持
//   V3 eIn 态 fIn=99 → eAbove（bAboveEdge 单拍）；fIn=94（< fHigh-fHyst）→ eIn
//   V4 fIn 跳变 -5 → 105：eBelow 一步直达 eAbove（单拍 bAboveEdge）
//   V5 fLow >= fHigh → eCfg + eZone = eIn；fIn = NaN → eInput + eZone = eIn
//   V6 bEn = FALSE → eZone = eIn、全出口清零（R303）
//   V7 非法枚举态（强改 _eZone）→ ELSE 兜底回 eIn + eCfg
// 修订记录 Revision  :
//   2026-11-22  v1.0.0  R65 首版（批 2 · 序号 6）
// ==============================================================================
TYPE E_DL_HbmZone :
(
    eBelow := 0,  // 下带：fIn 低于下带界 / below, the input under the lower band edge
    eIn    := 10, // 中带：fIn 在带内（安全中位）/ inside, the safe middle zone
    eAbove := 20  // 上带：fIn 高于上带界 / above, the input over the upper band edge
);
END_TYPE

TYPE E_DL_HbmErr :
(
    eNone  := 0,  // 无错 / no error
    eCfg   := 10, // 组态非法（fLow / fHigh / fHyst 域非法）/ an illegal configuration
    eInput := 20  // 输入非有限（fIn 为 NaN / Inf / 超幅值）/ a non finite input
);
END_TYPE

FUNCTION_BLOCK FB_DL_HysteresisBandMon
VAR_INPUT
    fIn   : LREAL;               // 监视输入 [工程单位] / the monitored input
    fLow  : LREAL := 0.0;        // 区间下界 [工程单位]，须 < fHigh / the lower band edge
    fHigh : LREAL := 100.0;      // 区间上界 [工程单位]，须 > fLow / the upper band edge
    fHyst : LREAL := 0.0;        // 迟滞半带宽 [工程单位]，须 [0, fHigh - fLow) / the hysteresis half band
    bEn   : BOOL := TRUE;        // 使能 [-]，FALSE 时出口清零回中位（R303）/ the enable
END_VAR
VAR_OUTPUT
    eZone      : E_DL_HbmZone := E_DL_HbmZone.eIn; // 区间状态出口 [状态]（安全中位初值）/ the zone outlet, safe middle initial
    bBelowEdge : BOOL := FALSE;  // 进入下带沿脉冲 [-]，单拍有效 / the below entry edge pulse, single scan
    bAboveEdge : BOOL := FALSE;  // 进入上带沿脉冲 [-]，单拍有效 / the above entry edge pulse, single scan
    bErr       : BOOL := FALSE;  // 错误标志 [-]，eCfg / eInput 置位 / the error flag
    eErr       : E_DL_HbmErr := E_DL_HbmErr.eNone; // 错误码出口 [码] / the error code outlet
END_VAR
VAR
    _eZone     : E_DL_HbmZone := E_DL_HbmZone.eIn; // 内部状态寄存器 [状态] / the internal state register
    _eZonePrev : E_DL_HbmZone := E_DL_HbmZone.eIn; // 本拍前态快照 [状态]（沿判定基准）/ the previous zone snapshot, the edge baseline
    _bCfgBad   : BOOL;           // 组态非法标志（逐拍重算）/ the configuration fault flag
    _bInBad    : BOOL;           // 输入非有限标志（逐拍重算）/ the input fault flag
END_VAR
VAR CONSTANT
    DL_HBM_FMAX : LREAL := 1.0E30; // 非有限筛查幅值上限 [工程单位] / the finiteness screening cap
END_VAR

// 段 1｜单拍沿脉冲与错误出口预清零（R256 统一出口预置）/ segment 1, the single scan preset
bBelowEdge := FALSE;             // 下带沿脉冲预清零 / preset the below edge false
bAboveEdge := FALSE;             // 上带沿脉冲预清零 / preset the above edge false
bErr       := FALSE;             // 错误标志预清零 / preset the error flag false
eErr       := E_DL_HbmErr.eNone; // 错误码预置无错 / preset the code to none

// 段 2｜失能分支：出口清零回安全中位，不置错（R303 离相清零声明行）/ segment 2, the disabled branch
IF NOT bEn THEN                  // 失能 / disabled
    _eZone := E_DL_HbmZone.eIn;  // 强制安全中位 / force the safe middle
    eZone := _eZone;             // 状态出口 / the zone outlet
    bBelowEdge := FALSE;         // 沿脉冲清零 / clear the below edge
    bAboveEdge := FALSE;         // 沿脉冲清零 / clear the above edge
    bErr := FALSE;               // 失能不是故障 / a disabled device is not a fault
    eErr := E_DL_HbmErr.eNone;   // 失能不发码 / no code while disabled
    RETURN;                      // 早退 / early return
END_IF

// 段 3｜组态守卫（边界一：四判据逐项点名，R272）/ segment 3, the configuration guard
_bCfgBad := (fLow >= fHigh)                                  // 下界不低于上界 / the lower edge not under the upper
         OR (fHyst < 0.0)                                    // 迟滞为负 / a negative hysteresis
         OR (fHyst >= (fHigh - fLow))                        // 迟滞吞没整带 / the hysteresis swallowing the whole band
         OR (fLow <> fLow) OR ((fLow - fLow) <> 0.0) OR (ABS(fLow) > DL_HBM_FMAX)      // fLow 非有限 / fLow non finite
         OR (fHigh <> fHigh) OR ((fHigh - fHigh) <> 0.0) OR (ABS(fHigh) > DL_HBM_FMAX) // fHigh 非有限 / fHigh non finite
         OR (fHyst <> fHyst) OR ((fHyst - fHyst) <> 0.0) OR (ABS(fHyst) > DL_HBM_FMAX); // fHyst 非有限 / fHyst non finite
IF _bCfgBad THEN                 // 组态非法 / an illegal configuration
    _eZone := E_DL_HbmZone.eIn;  // 强制安全中位（边界一）/ force the safe middle
    eZone := _eZone;             // 状态出口 / the zone outlet
    bErr := TRUE;                // 错误标志置位 / raise the error flag
    eErr := E_DL_HbmErr.eCfg;    // 信息级 0747：组态非法 / the configuration code
    RETURN;                      // 早退（沿脉冲保持段 1 预清零）/ early return
END_IF

// 段 4｜输入守卫（边界二：NaN 自反判 + Inf 差值自反判 + 幅值上界）/ segment 4, the input guard
_bInBad := (fIn <> fIn) OR ((fIn - fIn) <> 0.0) OR (ABS(fIn) > DL_HBM_FMAX); // 输入非有限 / the input non finite
IF _bInBad THEN                  // 输入无效 / an invalid input
    _eZone := E_DL_HbmZone.eIn;  // 强制安全中位（边界二）/ force the safe middle
    eZone := _eZone;             // 状态出口 / the zone outlet
    bErr := TRUE;                // 错误标志置位 / raise the error flag
    eErr := E_DL_HbmErr.eInput;  // 信息级 0748：输入非有限 / the input code
    RETURN;                      // 早退（沿脉冲保持段 1 预清零）/ early return
END_IF

// 段 5｜三带状态机（ENUM + CASE + ELSE 兜底，边界三 / 六）/ segment 5, the three zone machine
_eZonePrev := _eZone;            // 本拍前态快照（沿判定基准，边界四）/ snapshot the previous zone
CASE _eZone OF
    E_DL_HbmZone.eBelow:         // 下带 / the below zone
        IF fIn > fHigh THEN      // 跨带跳变直达上界之上（边界三一步直达）/ a jump beyond the upper edge
            _eZone := E_DL_HbmZone.eAbove; // 一步迁入上带 / straight to the above zone
        ELSIF fIn > (fLow + fHyst) THEN // 越过下带迟滞恢复线 / over the lower recovery line
            _eZone := E_DL_HbmZone.eIn;    // 迁入中带 / enter the inside zone
        END_IF
    E_DL_HbmZone.eIn:            // 中带 / the inside zone
        IF fIn < fLow THEN       // 跌破下界（严格小于，边界三）/ under the lower edge
            _eZone := E_DL_HbmZone.eBelow; // 迁入下带 / enter the below zone
        ELSIF fIn > fHigh THEN   // 越过上界（严格大于）/ over the upper edge
            _eZone := E_DL_HbmZone.eAbove; // 迁入上带 / enter the above zone
        END_IF
    E_DL_HbmZone.eAbove:         // 上带 / the above zone
        IF fIn < fLow THEN       // 跨带跳变跌破下界 / a jump under the lower edge
            _eZone := E_DL_HbmZone.eBelow; // 一步迁入下带 / straight to the below zone
        ELSIF fIn < (fHigh - fHyst) THEN // 跌破上带迟滞恢复线 / under the upper recovery line
            _eZone := E_DL_HbmZone.eIn;    // 迁入中带 / enter the inside zone
        END_IF
    ELSE                         // 非法枚举值拦截（边界六：回中位 + 组态族合并码，R90 反证句见码表）/ the illegal enumeration guard
        _eZone := E_DL_HbmZone.eIn; // 强制回安全中位 / force back to the safe middle
        bErr := TRUE;            // 错误标志置位（禁静默）/ raise the error flag
        eErr := E_DL_HbmErr.eCfg; // 归并组态族一码（出口同形不可区分，R90）/ merged into the configuration code
END_CASE

// 段 6｜沿脉冲与状态出口（边界四：基准 = 本拍前态快照，单拍有效）/ segment 6, the edges and the zone outlet
bBelowEdge := (_eZone = E_DL_HbmZone.eBelow) AND (_eZonePrev <> E_DL_HbmZone.eBelow); // 进入下带沿 / the below entry edge
bAboveEdge := (_eZone = E_DL_HbmZone.eAbove) AND (_eZonePrev <> E_DL_HbmZone.eAbove); // 进入上带沿 / the above entry edge
eZone := _eZone;                 // 状态出口（名实双出口同源，R191）/ the zone outlet
END_FUNCTION_BLOCK

(* ---- FB_DL_ImpulseRelay.st ---- *)
(*
  ==================================================================
  组件名 Component  : FB_DL_ImpulseRelay
  分类   Category   : DL_Base
  前缀   Naming     : FB_DL_ ｜ b/n/u/f/t/e 类型前缀制（R265）
  版本   Version    : 1.0.0
  功能   Purpose    : 沿触发定宽脉冲输出（按钮/点动 → 固定时长）：bTrig
                      上升沿置 bPulse，内部 tonPulse（PT = tPulseWidth）
                      定宽计时，计时到清 bPulse。重触发语义：脉宽运行中
                      再来沿，边沿拍强制 TON 计时基复位（IN 置 FALSE 一
                      拍，使 ET 归零重起）——重触发后的脉冲为完整新脉宽
                      （非残留余宽）。tPulseWidth ≤ T#0MS 配置非法电平
                      面码 01，故障拍不出脉冲。
  来源   Source     : t1-1-oscat-basic（定宽脉冲继电为 OSCAT 基础库公开
                      功能语义，clean-room 重写，零源码复制）
  互引   Cross-ref  : FB_DL_TpEx / FB_DL_PulseStretch（同族脉冲邻件：
                      TpEx 为脉宽可变触发延时变体，PulseStretch 为展宽
                      件，本件为固定脉宽沿触发口径属主）
  平台   Platform   : 纯 IEC 61131-3（R_TRIG/TON/TIME 比较）
  依赖   Depends    : 仅 Standard.library（R_TRIG/TON 属标准件）
  红线   Redline    : R1 零全局/VAR_EXTERNAL/R2 零 %I/%Q/R3 纯 IEC 标准
                      R4 配置闸显式 + TON/沿实例段 0 无条件刷新/R5 全变
                      量双语同行注释/R6 配置故障电平面无状态机（CASE 不
                      适用，头注说明）/R7 rtTrig/tonPulse 无条件周期调用
                      /R8 阈值常量化
  契约   Contract   : 码 01 配置非法为电平面（当拍复判）：故障拍 bPulse=
                      FALSE、bError=TRUE，恢复即恢复（恢复拍即触发沿则
                      照常出脉冲，同拍合法事件优先 R275）。bPulse 名实
                      双出口：bPulse=TRUE ⟺ tonPulse 计时窗内或边沿拍。
  错误码 Codes      : 01【故障级·电平面】tPulseWidth ≤ T#0MS 配置非法，
                      不出脉冲
  码位反证 Note     : 单码件（R90）：唯一失效面为脉宽配置面，无并置分立
                      依据；码 01 置 bError（故障级 3 行内配对，R45）。
  验收   Acceptance : V1 沿触发 → bPulse=TRUE 持续 tPulseWidth 后自落
                      ｜ V2 脉宽中途再沿 → 计时重起，总宽 ≈ 重触发时刻
                      + tPulseWidth ｜ V3 tPulseWidth=0 → 码 01（电平
                      面）｜ V4 连续 bTrig=TRUE → 仅首个沿出脉冲（沿触
                      发非电平触发）｜ V5 恢复合法脉宽 → 立即可触发
  变更   Revision   : 2026-11-22  v1.0.0  R67 首版（编码阶段批 3 序 4）
  ==================================================================
*)
FUNCTION_BLOCK FB_DL_ImpulseRelay
VAR_INPUT
    bTrig       : BOOL := FALSE;   // 触发输入（上升沿出脉冲）[-] / the trigger input, pulse on the rising edge
    tPulseWidth : TIME := T#1S;    // 脉宽 [ms]，须 > 0 / the pulse width, must be positive
END_VAR
VAR_OUTPUT
    bPulse   : BOOL := FALSE;       // 定宽脉冲输出 [-] / the fixed width pulse output
    bError   : BOOL := FALSE;       // 配置故障标志（电平面，恢复即清，R45 配对）/ the configuration fault flag
    uErrorId : UDINT := 16#0000_0000; // 错误码，0=正常，01 见头注 [码] / the error code [code]
END_VAR
VAR
    rtTrig   : R_TRIG;              // 触发沿实例，段 0 无条件刷新 / the trigger edge instance refreshed unconditionally
    tonPulse : TON;                 // 定宽计时实例，段 0 无条件刷新 / the width timer instance refreshed unconditionally
    _bCfgOk  : BOOL := FALSE;       // 本拍配置有效性 [-] / the per scan configuration validity
END_VAR
VAR CONSTANT
    IRL_ERR_NONE : UDINT := 16#0000_0000;  // 无错误 [码] / no error [code]
    IRL_ERR_CFG  : UDINT := 16#0000_0001;  // 码 01：脉宽配置非法 / code 01, illegal pulse width
END_VAR

(*------------------------------------------------------------------------------
 * 段 0｜沿检测与定时器无条件刷新区（红线 R7）：严禁移入 IF / CASE
 *      The edge and the timer refresh unconditionally, never inside a branch
 *-----------------------------------------------------------------------------*)
rtTrig(CLK := bTrig);                        // 触发沿 / the trigger edge
tonPulse(IN := bPulse AND NOT rtTrig.Q, PT := tPulseWidth);  // 定宽计时：边沿拍强制 IN=FALSE 使 ET 归零重起（重触发完整新脉宽，R188 自复位语义）/ the width timing, the edge scan resets the timing base

(*------------------------------------------------------------------------------
 * 段 1｜错误码本拍预置 + 配置闸（电平面，当拍复判，码 01）
 *      The error code preset and the configuration gate
 *-----------------------------------------------------------------------------*)
uErrorId := IRL_ERR_NONE;       // 预置无错误 / preset no error
_bCfgOk := (tPulseWidth > T#0MS);  // 配置闸（TIME 直接比较，三平台一致）/ the configuration gate
IF NOT _bCfgOk THEN
    bError := TRUE;             // 故障标志（R45 配对，故障级 3 行内置）/ the fault flag
    uErrorId := IRL_ERR_CFG;    // 码 01 / code 01
    bPulse := FALSE;            // 故障拍不出脉冲（安全缺省）/ no pulse on fault
    RETURN;                     // 结构早退（tonPulse 已刷，段 0 契约不破）/ structural early return
ELSE
    bError := FALSE;            // 配置恢复即清（电平面契约）/ cleared when the configuration recovers
END_IF

(*------------------------------------------------------------------------------
 * 段 2｜沿触发置位（同拍合法事件优先于计时窗判定，R275）
 *      The edge set, the legal event before the window verdict
 *-----------------------------------------------------------------------------*)
IF rtTrig.Q THEN
    bPulse := TRUE;             // 沿置脉冲 / set the pulse on the edge
END_IF

(*------------------------------------------------------------------------------
 * 段 3｜计时窗到清位（段 0 已刷 tonPulse：边沿拍 Q=FALSE 不误清，下拍起算）
 *      The window expiry clears the pulse, the edge scan never clears
 *-----------------------------------------------------------------------------*)
IF tonPulse.Q THEN
    bPulse := FALSE;            // 脉宽到落脉冲 / drop the pulse on expiry
END_IF
END_FUNCTION_BLOCK
